HMI tags "Default tag table"
   "7" : Bool = PLC "ป้อนรหัส Barcode" AT %I100.6, 1 s
   "Alarms_All" : Word = PLC "บันทึกผลการเคลื่อนที่ ไว้ที่ Excell_DB".Alarms AT %DB1.DBX0.0, 1 s
   "Barcode1" : Word = PLC Barcode1 AT %MW2000, 1 s
   "Barcode10" : Word = PLC Barcode10 AT %MW2018, 1 s
   "Barcode100" : Word = PLC Barcode100 AT %MW2198, 1 s
   "Barcode101" : Word = PLC Barcode101 AT %MW2200, 1 s
   "Barcode102" : Word = PLC Barcode102 AT %MW2202, 1 s
   "Barcode103" : Word = PLC Barcode103 AT %MW2204, 1 s
   "Barcode104" : Word = PLC Barcode104 AT %MW2206, 1 s
   "Barcode105" : Word = PLC Barcode105 AT %MW2208, 1 s
   "Barcode106" : Word = PLC Barcode106 AT %MW2210, 1 s
   "Barcode107" : Word = PLC Barcode107 AT %MW2212, 1 s
   "Barcode108" : Word = PLC Barcode108 AT %MW2214, 1 s
   "Barcode109" : Word = PLC Barcode109 AT %MW2216, 1 s
   "Barcode11" : Word = PLC Barcode11 AT %MW2020, 1 s
   "Barcode110" : Word = PLC Barcode110 AT %MW2218, 1 s
   "Barcode111" : Word = PLC Barcode111 AT %MW2220, 1 s
   "Barcode112" : Word = PLC Barcode112 AT %MW2222, 1 s
   "Barcode113" : Word = PLC Barcode113 AT %MW2224, 1 s
   "Barcode114" : Word = PLC Barcode114 AT %MW2226, 1 s
   "Barcode115" : Word = PLC Barcode115 AT %MW2228, 1 s
   "Barcode116" : Word = PLC Barcode116 AT %MW2230, 1 s
   "Barcode117" : Word = PLC Barcode117 AT %MW2232, 1 s
   "Barcode118" : Word = PLC Barcode118 AT %MW2234, 1 s
   "Barcode119" : Word = PLC Barcode119 AT %MW2236, 1 s
   "Barcode12" : Word = PLC Barcode12 AT %MW2022, 1 s
   "Barcode120" : Word = PLC Barcode120 AT %MW2238, 1 s
   "Barcode121" : Word = PLC Barcode121 AT %MW2240, 1 s
   "Barcode122" : Word = PLC Barcode122 AT %MW2242, 1 s
   "Barcode123" : Word = PLC Barcode123 AT %MW2244, 1 s
   "Barcode124" : Word = PLC Barcode124 AT %MW2246, 1 s
   "Barcode125" : Word = PLC Barcode125 AT %MW2248, 1 s
   "Barcode126" : Word = PLC Barcode126 AT %MW2250, 1 s
   "Barcode127" : Word = PLC Barcode127 AT %MW2252, 1 s
   "Barcode128" : Word = PLC Barcode128 AT %MW2254, 1 s
   "Barcode129" : Word = PLC Barcode129 AT %MW2256, 1 s
   "Barcode13" : Word = PLC Barcode13 AT %MW2024, 1 s
   "Barcode130" : Word = PLC Barcode130 AT %MW2258, 1 s
   "Barcode131" : Word = PLC Barcode131 AT %MW2260, 1 s
   "Barcode132" : Word = PLC Barcode132 AT %MW2262, 1 s
   "Barcode133" : Word = PLC Barcode133 AT %MW2264, 1 s
   "Barcode134" : Word = PLC Barcode134 AT %MW2266, 1 s
   "Barcode135" : Word = PLC Barcode135 AT %MW2268, 1 s
   "Barcode136" : Word = PLC Barcode136 AT %MW2270, 1 s
   "Barcode137" : Word = PLC Barcode137 AT %MW2272, 1 s
   "Barcode138" : Word = PLC Barcode138 AT %MW2274, 1 s
   "Barcode139" : Word = PLC Barcode139 AT %MW2276, 1 s
   "Barcode14" : Word = PLC Barcode14 AT %MW2026, 1 s
   "Barcode140" : Word = PLC Barcode140 AT %MW2278, 1 s
   "Barcode141" : Word = PLC Barcode141 AT %MW2280, 1 s
   "Barcode142" : Word = PLC Barcode142 AT %MW2282, 1 s
   "Barcode143" : Word = PLC Barcode143 AT %MW2284, 1 s
   "Barcode144" : Word = PLC Barcode144 AT %MW2286, 1 s
   "Barcode145" : Word = PLC Barcode145 AT %MW2288, 1 s
   "Barcode146" : Word = PLC Barcode146 AT %MW2290, 1 s
   "Barcode147" : Word = PLC Barcode147 AT %MW2292, 1 s
   "Barcode148" : Word = PLC Barcode148 AT %MW2294, 1 s
   "Barcode149" : Word = PLC Barcode149 AT %MW2296, 1 s
   "Barcode15" : Word = PLC Barcode15 AT %MW2028, 1 s
   "Barcode150" : Word = PLC Barcode150 AT %MW2298, 1 s
   "Barcode151" : Word = PLC Barcode151 AT %MW2300, 1 s
   "Barcode152" : Word = PLC Barcode152 AT %MW2302, 1 s
   "Barcode153" : Word = PLC Barcode153 AT %MW2304, 1 s
   "Barcode154" : Word = PLC Barcode154 AT %MW2306, 1 s
   "Barcode155" : Word = PLC Barcode155 AT %MW2308, 1 s
   "Barcode156" : Word = PLC Barcode156 AT %MW2310, 1 s
   "Barcode157" : Word = PLC Barcode157 AT %MW2312, 1 s
   "Barcode158" : Word = PLC Barcode158 AT %MW2314, 1 s
   "Barcode159" : Word = PLC Barcode159 AT %MW2316, 1 s
   "Barcode16" : Word = PLC Barcode16 AT %MW2030, 1 s
   "Barcode160" : Word = PLC Barcode160 AT %MW2318, 1 s
   "Barcode161" : Word = PLC Barcode161 AT %MW2320, 1 s
   "Barcode162" : Word = PLC Barcode162 AT %MW2322, 1 s
   "Barcode163" : Word = PLC Barcode163 AT %MW2324, 1 s
   "Barcode164" : Word = PLC Barcode164 AT %MW2326, 1 s
   "Barcode165" : Word = PLC Barcode165 AT %MW2328, 1 s
   "Barcode166" : Word = PLC Barcode166 AT %MW2330, 1 s
   "Barcode167" : Word = PLC Barcode167 AT %MW2332, 1 s
   "Barcode168" : Word = PLC Barcode168 AT %MW2334, 1 s
   "Barcode169" : Word = PLC Barcode169 AT %MW2336, 1 s
   "Barcode17" : Word = PLC Barcode17 AT %MW2032, 1 s
   "Barcode170" : Word = PLC Barcode170 AT %MW2338, 1 s
   "Barcode171" : Word = PLC Barcode171 AT %MW2340, 1 s
   "Barcode172" : Word = PLC Barcode172 AT %MW2342, 1 s
   "Barcode173" : Word = PLC Barcode173 AT %MW2344, 1 s
   "Barcode174" : Word = PLC Barcode174 AT %MW2346, 1 s
   "Barcode175" : Word = PLC Barcode175 AT %MW2348, 1 s
   "Barcode176" : Word = PLC Barcode176 AT %MW2350, 1 s
   "Barcode177" : Word = PLC Barcode177 AT %MW2352, 1 s
   "Barcode178" : Word = PLC Barcode178 AT %MW2354, 1 s
   "Barcode179" : Word = PLC Barcode179 AT %MW2356, 1 s
   "Barcode18" : Word = PLC Barcode18 AT %MW2034, 1 s
   "Barcode180" : Word = PLC Barcode180 AT %MW2358, 1 s
   "Barcode181" : Word = PLC Barcode181 AT %MW2360, 1 s
   "Barcode182" : Word = PLC Barcode182 AT %MW2362, 1 s
   "Barcode183" : Word = PLC Barcode183 AT %MW2364, 1 s
   "Barcode184" : Word = PLC Barcode184 AT %MW2366, 1 s
   "Barcode185" : Word = PLC Barcode185 AT %MW2368, 1 s
   "Barcode186" : Word = PLC Barcode186 AT %MW2370, 1 s
   "Barcode187" : Word = PLC Barcode187 AT %MW2372, 1 s
   "Barcode188" : Word = PLC Barcode188 AT %MW2374, 1 s
   "Barcode189" : Word = PLC Barcode189 AT %MW2376, 1 s
   "Barcode19" : Word = PLC Barcode19 AT %MW2036, 1 s
   "Barcode190" : Word = PLC Barcode190 AT %MW2378, 1 s
   "Barcode191" : Word = PLC Barcode191 AT %MW2380, 1 s
   "Barcode192" : Word = PLC Barcode192 AT %MW2382, 1 s
   "Barcode193" : Word = PLC Barcode193 AT %MW2384, 1 s
   "Barcode194" : Word = PLC Barcode194 AT %MW2386, 1 s
   "Barcode195" : Word = PLC Barcode195 AT %MW2388, 1 s
   "Barcode196" : Word = PLC Barcode196 AT %MW2390, 1 s
   "Barcode197" : Word = PLC Barcode197 AT %MW2392, 1 s
   "Barcode198" : Word = PLC Barcode198 AT %MW2394, 1 s
   "Barcode199" : Word = PLC Barcode199 AT %MW2396, 1 s
   "Barcode2" : Word = PLC Barcode2 AT %MW2002, 1 s
   "Barcode20" : Word = PLC Barcode20 AT %MW2038, 1 s
   "Barcode200" : Word = PLC Barcode200 AT %MW2398, 1 s
   "Barcode201" : Word = PLC Barcode201 AT %MW2400, 1 s
   "Barcode202" : Word = PLC Barcode202 AT %MW2402, 1 s
   "Barcode203" : Word = PLC Barcode203 AT %MW2404, 1 s
   "Barcode204" : Word = PLC Barcode204 AT %MW2406, 1 s
   "Barcode205" : Word = PLC Barcode205 AT %MW2408, 1 s
   "Barcode206" : Word = PLC Barcode206 AT %MW2410, 1 s
   "Barcode207" : Word = PLC Barcode207 AT %MW2412, 1 s
   "Barcode208" : Word = PLC Barcode208 AT %MW2414, 1 s
   "Barcode209" : Word = PLC Barcode209 AT %MW2416, 1 s
   "Barcode21" : Word = PLC Barcode21 AT %MW2040, 1 s
   "Barcode210" : Word = PLC Barcode210 AT %MW2418, 1 s
   "Barcode211" : Word = PLC Barcode211 AT %MW2420, 1 s
   "Barcode212" : Word = PLC Barcode212 AT %MW2422, 1 s
   "Barcode213" : Word = PLC Barcode213 AT %MW2424, 1 s
   "Barcode214" : Word = PLC Barcode214 AT %MW2426, 1 s
   "Barcode215" : Word = PLC Barcode215 AT %MW2428, 1 s
   "Barcode216" : Word = PLC Barcode216 AT %MW2430, 1 s
   "Barcode217" : Word = PLC Barcode217 AT %MW2432, 1 s
   "Barcode218" : Word = PLC Barcode218 AT %MW2434, 1 s
   "Barcode219" : Word = PLC Barcode219 AT %MW2436, 1 s
   "Barcode22" : Word = PLC Barcode22 AT %MW2042, 1 s
   "Barcode220" : Word = PLC Barcode220 AT %MW2438, 1 s
   "Barcode221" : Word = PLC Barcode221 AT %MW2440, 1 s
   "Barcode222" : Word = PLC Barcode222 AT %MW2442, 1 s
   "Barcode223" : Word = PLC Barcode223 AT %MW2444, 1 s
   "Barcode224" : Word = PLC Barcode224 AT %MW2446, 1 s
   "Barcode225" : Word = PLC Barcode225 AT %MW2448, 1 s
   "Barcode226" : Word = PLC Barcode226 AT %MW2450, 1 s
   "Barcode227" : Word = PLC Barcode227 AT %MW2452, 1 s
   "Barcode228" : Word = PLC Barcode228 AT %MW2454, 1 s
   "Barcode229" : Word = PLC Barcode229 AT %MW2456, 1 s
   "Barcode23" : Word = PLC Barcode23 AT %MW2044, 1 s
   "Barcode230" : Word = PLC Barcode230 AT %MW2458, 1 s
   "Barcode231" : Word = PLC Barcode231 AT %MW2460, 1 s
   "Barcode232" : Word = PLC Barcode232 AT %MW2462, 1 s
   "Barcode233" : Word = PLC Barcode233 AT %MW2464, 1 s
   "Barcode234" : Word = PLC Barcode234 AT %MW2466, 1 s
   "Barcode235" : Word = PLC Barcode235 AT %MW2468, 1 s
   "Barcode236" : Word = PLC Barcode236 AT %MW2470, 1 s
   "Barcode237" : Word = PLC Barcode237 AT %MW2472, 1 s
   "Barcode238" : Word = PLC Barcode238 AT %MW2474, 1 s
   "Barcode239" : Word = PLC Barcode239 AT %MW2476, 1 s
   "Barcode24" : Word = PLC Barcode24 AT %MW2046, 1 s
   "Barcode240" : Word = PLC Barcode240 AT %MW2478, 1 s
   "Barcode241" : Word = PLC Barcode241 AT %MW2480, 1 s
   "Barcode242" : Word = PLC Barcode242 AT %MW2482, 1 s
   "Barcode243" : Word = PLC Barcode243 AT %MW2484, 1 s
   "Barcode244" : Word = PLC Barcode244 AT %MW2486, 1 s
   "Barcode245" : Word = PLC Barcode245 AT %MW2488, 1 s
   "Barcode246" : Word = PLC Barcode246 AT %MW2490, 1 s
   "Barcode247" : Word = PLC Barcode247 AT %MW2492, 1 s
   "Barcode248" : Word = PLC Barcode248 AT %MW2494, 1 s
   "Barcode249" : Word = PLC Barcode249 AT %MW2496, 1 s
   "Barcode25" : Word = PLC Barcode25 AT %MW2048, 1 s
   "Barcode250" : Word = PLC Barcode250 AT %MW2498, 1 s
   "Barcode251" : Word = PLC Barcode251 AT %MW2500, 1 s
   "Barcode252" : Word = PLC Barcode252 AT %MW2502, 1 s
   "Barcode253" : Word = PLC Barcode253 AT %MW2504, 1 s
   "Barcode254" : Word = PLC Barcode254 AT %MW2506, 1 s
   "Barcode255" : Word = PLC Barcode255 AT %MW2508, 1 s
   "Barcode256" : Word = PLC Barcode256 AT %MW2510, 1 s
   "Barcode257" : Word = PLC Barcode257 AT %MW2512, 1 s
   "Barcode258" : Word = PLC Barcode258 AT %MW2514, 1 s
   "Barcode259" : Word = PLC Barcode259 AT %MW2516, 1 s
   "Barcode26" : Word = PLC Barcode26 AT %MW2050, 1 s
   "Barcode260" : Word = PLC Barcode260 AT %MW2518, 1 s
   "Barcode261" : Word = PLC Barcode261 AT %MW2520, 1 s
   "Barcode262" : Word = PLC Barcode262 AT %MW2522, 1 s
   "Barcode263" : Word = PLC Barcode263 AT %MW2524, 1 s
   "Barcode264" : Word = PLC Barcode264 AT %MW2526, 1 s
   "Barcode265" : Word = PLC Barcode265 AT %MW2528, 1 s
   "Barcode266" : Word = PLC Barcode266 AT %MW2530, 1 s
   "Barcode267" : Word = PLC Barcode267 AT %MW2532, 1 s
   "Barcode268" : Word = PLC Barcode268 AT %MW2534, 1 s
   "Barcode269" : Word = PLC Barcode269 AT %MW2536, 1 s
   "Barcode27" : Word = PLC Barcode27 AT %MW2052, 1 s
   "Barcode270" : Word = PLC Barcode270 AT %MW2538, 1 s
   "Barcode271" : Word = PLC Barcode271 AT %MW2540, 1 s
   "Barcode272" : Word = PLC Barcode272 AT %MW2542, 1 s
   "Barcode273" : Word = PLC Barcode273 AT %MW2544, 1 s
   "Barcode274" : Word = PLC Barcode274 AT %MW2546, 1 s
   "Barcode275" : Word = PLC Barcode275 AT %MW2548, 1 s
   "Barcode276" : Word = PLC Barcode276 AT %MW2550, 1 s
   "Barcode277" : Word = PLC Barcode277 AT %MW2552, 1 s
   "Barcode278" : Word = PLC Barcode278 AT %MW2554, 1 s
   "Barcode279" : Word = PLC Barcode279 AT %MW2556, 1 s
   "Barcode28" : Word = PLC Barcode28 AT %MW2054, 1 s
   "Barcode280" : Word = PLC Barcode280 AT %MW2558, 1 s
   "Barcode281" : Word = PLC Barcode281 AT %MW2560, 1 s
   "Barcode282" : Word = PLC Barcode282 AT %MW2562, 1 s
   "Barcode283" : Word = PLC Barcode283 AT %MW2564, 1 s
   "Barcode284" : Word = PLC Barcode284 AT %MW2566, 1 s
   "Barcode285" : Word = PLC Barcode285 AT %MW2568, 1 s
   "Barcode286" : Word = PLC Barcode286 AT %MW2570, 1 s
   "Barcode287" : Word = PLC Barcode287 AT %MW2572, 1 s
   "Barcode288" : Word = PLC Barcode288 AT %MW2574, 1 s
   "Barcode289" : Word = PLC Barcode289 AT %MW2576, 1 s
   "Barcode29" : Word = PLC Barcode29 AT %MW2056, 1 s
   "Barcode290" : Word = PLC Barcode290 AT %MW2578, 1 s
   "Barcode291" : Word = PLC Barcode291 AT %MW2580, 1 s
   "Barcode292" : Word = PLC Barcode292 AT %MW2582, 1 s
   "Barcode293" : Word = PLC Barcode293 AT %MW2584, 1 s
   "Barcode294" : Word = PLC Barcode294 AT %MW2586, 1 s
   "Barcode295" : Word = PLC Barcode295 AT %MW2588, 1 s
   "Barcode296" : Word = PLC Barcode296 AT %MW2590, 1 s
   "Barcode297" : Word = PLC Barcode297 AT %MW2592, 1 s
   "Barcode298" : Word = PLC Barcode298 AT %MW2594, 1 s
   "Barcode299" : Word = PLC Barcode299 AT %MW2596, 1 s
   "Barcode3" : Word = PLC Barcode3 AT %MW2004, 1 s
   "Barcode30" : Word = PLC Barcode30 AT %MW2058, 1 s
   "Barcode300" : Word = PLC Barcode300 AT %MW2598, 1 s
   "Barcode301" : Word = PLC Barcode301 AT %MW2600, 1 s
   "Barcode302" : Word = PLC Barcode302 AT %MW2602, 1 s
   "Barcode303" : Word = PLC Barcode303 AT %MW2604, 1 s
   "Barcode304" : Word = PLC Barcode304 AT %MW2606, 1 s
   "Barcode305" : Word = PLC Barcode305 AT %MW2608, 1 s
   "Barcode306" : Word = PLC Barcode306 AT %MW2610, 1 s
   "Barcode307" : Word = PLC Barcode307 AT %MW2612, 1 s
   "Barcode308" : Word = PLC Barcode308 AT %MW2614, 1 s
   "Barcode309" : Word = PLC Barcode309 AT %MW2616, 1 s
   "Barcode31" : Word = PLC Barcode31 AT %MW2060, 1 s
   "Barcode310" : Word = PLC Barcode310 AT %MW2618, 1 s
   "Barcode311" : Word = PLC Barcode311 AT %MW2620, 1 s
   "Barcode312" : Word = PLC Barcode312 AT %MW2622, 1 s
   "Barcode313" : Word = PLC Barcode313 AT %MW2624, 1 s
   "Barcode314" : Word = PLC Barcode314 AT %MW2626, 1 s
   "Barcode315" : Word = PLC Barcode315 AT %MW2628, 1 s
   "Barcode316" : Word = PLC Barcode316 AT %MW2630, 1 s
   "Barcode317" : Word = PLC Barcode317 AT %MW2632, 1 s
   "Barcode318" : Word = PLC Barcode318 AT %MW2634, 1 s
   "Barcode319" : Word = PLC Barcode319 AT %MW2636, 1 s
   "Barcode32" : Word = PLC Barcode32 AT %MW2062, 1 s
   "Barcode320" : Word = PLC Barcode320 AT %MW2638, 1 s
   "Barcode321" : Word = PLC Barcode321 AT %MW2640, 1 s
   "Barcode322" : Word = PLC Barcode322 AT %MW2642, 1 s
   "Barcode323" : Word = PLC Barcode323 AT %MW2644, 1 s
   "Barcode324" : Word = PLC Barcode324 AT %MW2646, 1 s
   "Barcode325" : Word = PLC Barcode325 AT %MW2648, 1 s
   "Barcode326" : Word = PLC Barcode326 AT %MW2650, 1 s
   "Barcode327" : Word = PLC Barcode327 AT %MW2652, 1 s
   "Barcode328" : Word = PLC Barcode328 AT %MW2654, 1 s
   "Barcode329" : Word = PLC Barcode329 AT %MW2656, 1 s
   "Barcode33" : Word = PLC Barcode33 AT %MW2064, 1 s
   "Barcode330" : Word = PLC Barcode330 AT %MW2658, 1 s
   "Barcode331" : Word = PLC Barcode331 AT %MW2660, 1 s
   "Barcode332" : Word = PLC Barcode332 AT %MW2662, 1 s
   "Barcode333" : Word = PLC Barcode333 AT %MW2664, 1 s
   "Barcode334" : Word = PLC Barcode334 AT %MW2666, 1 s
   "Barcode335" : Word = PLC Barcode335 AT %MW2668, 1 s
   "Barcode336" : Word = PLC Barcode336 AT %MW2670, 1 s
   "Barcode337" : Word = PLC Barcode337 AT %MW2672, 1 s
   "Barcode338" : Word = PLC Barcode338 AT %MW2674, 1 s
   "Barcode339" : Word = PLC Barcode339 AT %MW2676, 1 s
   "Barcode34" : Word = PLC Barcode34 AT %MW2066, 1 s
   "Barcode340" : Word = PLC Barcode340 AT %MW2678, 1 s
   "Barcode341" : Word = PLC Barcode341 AT %MW2680, 1 s
   "Barcode342" : Word = PLC Barcode342 AT %MW2682, 1 s
   "Barcode343" : Word = PLC Barcode343 AT %MW2684, 1 s
   "Barcode344" : Word = PLC Barcode344 AT %MW2686, 1 s
   "Barcode345" : Word = PLC Barcode345 AT %MW2688, 1 s
   "Barcode346" : Word = PLC Barcode346 AT %MW2690, 1 s
   "Barcode347" : Word = PLC Barcode347 AT %MW2692, 1 s
   "Barcode348" : Word = PLC Barcode348 AT %MW2694, 1 s
   "Barcode349" : Word = PLC Barcode349 AT %MW2696, 1 s
   "Barcode35" : Word = PLC Barcode35 AT %MW2068, 1 s
   "Barcode350" : Word = PLC Barcode350 AT %MW2698, 1 s
   "Barcode351" : Word = PLC Barcode351 AT %MW2700, 1 s
   "Barcode352" : Word = PLC Barcode352 AT %MW2702, 1 s
   "Barcode353" : Word = PLC Barcode353 AT %MW2704, 1 s
   "Barcode354" : Word = PLC Barcode354 AT %MW2706, 1 s
   "Barcode355" : Word = PLC Barcode355 AT %MW2708, 1 s
   "Barcode356" : Word = PLC Barcode356 AT %MW2710, 1 s
   "Barcode357" : Word = PLC Barcode357 AT %MW2712, 1 s
   "Barcode358" : Word = PLC Barcode358 AT %MW2714, 1 s
   "Barcode359" : Word = PLC Barcode359 AT %MW2716, 1 s
   "Barcode36" : Word = PLC Barcode36 AT %MW2070, 1 s
   "Barcode360" : Word = PLC Barcode360 AT %MW2718, 1 s
   "Barcode361" : Word = PLC Barcode361 AT %MW2720, 1 s
   "Barcode362" : Word = PLC Barcode362 AT %MW2722, 1 s
   "Barcode363" : Word = PLC Barcode363 AT %MW2724, 1 s
   "Barcode364" : Word = PLC Barcode364 AT %MW2726, 1 s
   "Barcode365" : Word = PLC Barcode365 AT %MW2728, 1 s
   "Barcode366" : Word = PLC Barcode366 AT %MW2730, 1 s
   "Barcode367" : Word = PLC Barcode367 AT %MW2732, 1 s
   "Barcode368" : Word = PLC Barcode368 AT %MW2734, 1 s
   "Barcode369" : Word = PLC Barcode369 AT %MW2736, 1 s
   "Barcode37" : Word = PLC Barcode37 AT %MW2072, 1 s
   "Barcode370" : Word = PLC Barcode370 AT %MW2738, 1 s
   "Barcode371" : Word = PLC Barcode371 AT %MW2740, 1 s
   "Barcode372" : Word = PLC Barcode372 AT %MW2742, 1 s
   "Barcode373" : Word = PLC Barcode373 AT %MW2744, 1 s
   "Barcode374" : Word = PLC Barcode374 AT %MW2746, 1 s
   "Barcode375" : Word = PLC Barcode375 AT %MW2748, 1 s
   "Barcode376" : Word = PLC Barcode376 AT %MW2750, 1 s
   "Barcode377" : Word = PLC Barcode377 AT %MW2752, 1 s
   "Barcode378" : Word = PLC Barcode378 AT %MW2754, 1 s
   "Barcode379" : Word = PLC Barcode379 AT %MW2756, 1 s
   "Barcode38" : Word = PLC Barcode38 AT %MW2074, 1 s
   "Barcode380" : Word = PLC Barcode380 AT %MW2758, 1 s
   "Barcode381" : Word = PLC Barcode381 AT %MW2760, 1 s
   "Barcode382" : Word = PLC Barcode382 AT %MW2762, 1 s
   "Barcode383" : Word = PLC Barcode383 AT %MW2764, 1 s
   "Barcode384" : Word = PLC Barcode384 AT %MW2766, 1 s
   "Barcode385" : Word = PLC Barcode385 AT %MW2768, 1 s
   "Barcode386" : Word = PLC Barcode386 AT %MW2770, 1 s
   "Barcode387" : Word = PLC Barcode387 AT %MW2772, 1 s
   "Barcode388" : Word = PLC Barcode388 AT %MW2774, 1 s
   "Barcode389" : Word = PLC Barcode389 AT %MW2776, 1 s
   "Barcode39" : Word = PLC Barcode39 AT %MW2076, 1 s
   "Barcode390" : Word = PLC Barcode390 AT %MW2778, 1 s
   "Barcode391" : Word = PLC Barcode391 AT %MW2780, 1 s
   "Barcode392" : Word = PLC Barcode392 AT %MW2782, 1 s
   "Barcode393" : Word = PLC Barcode393 AT %MW2784, 1 s
   "Barcode394" : Word = PLC Barcode394 AT %MW2786, 1 s
   "Barcode395" : Word = PLC Barcode395 AT %MW2788, 1 s
   "Barcode396" : Word = PLC Barcode396 AT %MW2790, 1 s
   "Barcode397" : Word = PLC Barcode397 AT %MW2792, 1 s
   "Barcode398" : Word = PLC Barcode398 AT %MW2794, 1 s
   "Barcode399" : Word = PLC Barcode399 AT %MW2796, 1 s
   "Barcode4" : Word = PLC Barcode4 AT %MW2006, 1 s
   "Barcode40" : Word = PLC Barcode40 AT %MW2078, 1 s
   "Barcode400" : Word = PLC Barcode400 AT %MW2798, 1 s
   "Barcode401" : Word = PLC Barcode401 AT %MW2800, 1 s
   "Barcode402" : Word = PLC Barcode402 AT %MW2802, 1 s
   "Barcode403" : Word = PLC Barcode403 AT %MW2804, 1 s
   "Barcode404" : Word = PLC Barcode404 AT %MW2806, 1 s
   "Barcode405" : Word = PLC Barcode405 AT %MW2808, 1 s
   "Barcode406" : Word = PLC Barcode406 AT %MW2810, 1 s
   "Barcode407" : Word = PLC Barcode407 AT %MW2812, 1 s
   "Barcode408" : Word = PLC Barcode408 AT %MW2814, 1 s
   "Barcode409" : Word = PLC Barcode409 AT %MW2816, 1 s
   "Barcode41" : Word = PLC Barcode41 AT %MW2080, 1 s
   "Barcode410" : Word = PLC Barcode410 AT %MW2818, 1 s
   "Barcode411" : Word = PLC Barcode411 AT %MW2820, 1 s
   "Barcode412" : Word = PLC Barcode412 AT %MW2822, 1 s
   "Barcode413" : Word = PLC Barcode413 AT %MW2824, 1 s
   "Barcode414" : Word = PLC Barcode414 AT %MW2826, 1 s
   "Barcode415" : Word = PLC Barcode415 AT %MW2828, 1 s
   "Barcode416" : Word = PLC Barcode416 AT %MW2830, 1 s
   "Barcode417" : Word = PLC Barcode417 AT %MW2832, 1 s
   "Barcode418" : Word = PLC Barcode418 AT %MW2834, 1 s
   "Barcode419" : Word = PLC Barcode419 AT %MW2836, 1 s
   "Barcode42" : Word = PLC Barcode42 AT %MW2082, 1 s
   "Barcode420" : Word = PLC Barcode420 AT %MW2838, 1 s
   "Barcode421" : Word = PLC Barcode421 AT %MW2840, 1 s
   "Barcode422" : Word = PLC Barcode422 AT %MW2842, 1 s
   "Barcode423" : Word = PLC Barcode423 AT %MW2844, 1 s
   "Barcode424" : Word = PLC Barcode424 AT %MW2846, 1 s
   "Barcode425" : Word = PLC Barcode425 AT %MW2848, 1 s
   "Barcode426" : Word = PLC Barcode426 AT %MW2850, 1 s
   "Barcode427" : Word = PLC Barcode427 AT %MW2852, 1 s
   "Barcode428" : Word = PLC Barcode428 AT %MW2854, 1 s
   "Barcode429" : Word = PLC Barcode429 AT %MW2856, 1 s
   "Barcode43" : Word = PLC Barcode43 AT %MW2084, 1 s
   "Barcode430" : Word = PLC Barcode430 AT %MW2858, 1 s
   "Barcode431" : Word = PLC Barcode431 AT %MW2860, 1 s
   "Barcode432" : Word = PLC Barcode432 AT %MW2862, 1 s
   "Barcode433" : Word = PLC Barcode433 AT %MW2864, 1 s
   "Barcode434" : Word = PLC Barcode434 AT %MW2866, 1 s
   "Barcode435" : Word = PLC Barcode435 AT %MW2868, 1 s
   "Barcode436" : Word = PLC Barcode436 AT %MW2870, 1 s
   "Barcode437" : Word = PLC Barcode437 AT %MW2872, 1 s
   "Barcode438" : Word = PLC Barcode438 AT %MW2874, 1 s
   "Barcode439" : Word = PLC Barcode439 AT %MW2876, 1 s
   "Barcode44" : Word = PLC Barcode44 AT %MW2086, 1 s
   "Barcode440" : Word = PLC Barcode440 AT %MW2878, 1 s
   "Barcode441" : Word = PLC Barcode441 AT %MW2880, 1 s
   "Barcode442" : Word = PLC Barcode442 AT %MW2882, 1 s
   "Barcode443" : Word = PLC Barcode443 AT %MW2884, 1 s
   "Barcode444" : Word = PLC Barcode444 AT %MW2886, 1 s
   "Barcode445" : Word = PLC Barcode445 AT %MW2888, 1 s
   "Barcode446" : Word = PLC Barcode446 AT %MW2890, 1 s
   "Barcode447" : Word = PLC Barcode447 AT %MW2892, 1 s
   "Barcode448" : Word = PLC Barcode448 AT %MW2894, 1 s
   "Barcode449" : Word = PLC Barcode449 AT %MW2896, 1 s
   "Barcode45" : Word = PLC Barcode45 AT %MW2088, 1 s
   "Barcode450" : Word = PLC Barcode450 AT %MW2898, 1 s
   "Barcode451" : Word = PLC Barcode451 AT %MW2900, 1 s
   "Barcode452" : Word = PLC Barcode452 AT %MW2902, 1 s
   "Barcode453" : Word = PLC Barcode453 AT %MW2904, 1 s
   "Barcode454" : Word = PLC Barcode454 AT %MW2906, 1 s
   "Barcode455" : Word = PLC Barcode455 AT %MW2908, 1 s
   "Barcode456" : Word = PLC Barcode456 AT %MW2910, 1 s
   "Barcode457" : Word = PLC Barcode457 AT %MW2912, 1 s
   "Barcode458" : Word = PLC Barcode458 AT %MW2914, 1 s
   "Barcode459" : Word = PLC Barcode459 AT %MW2916, 1 s
   "Barcode46" : Word = PLC Barcode46 AT %MW2090, 1 s
   "Barcode460" : Word = PLC Barcode460 AT %MW2918, 1 s
   "Barcode461" : Word = PLC Barcode461 AT %MW2920, 1 s
   "Barcode462" : Word = PLC Barcode462 AT %MW2922, 1 s
   "Barcode463" : Word = PLC Barcode463 AT %MW2924, 1 s
   "Barcode464" : Word = PLC Barcode464 AT %MW2926, 1 s
   "Barcode465" : Word = PLC Barcode465 AT %MW2928, 1 s
   "Barcode466" : Word = PLC Barcode466 AT %MW2930, 1 s
   "Barcode467" : Word = PLC Barcode467 AT %MW2932, 1 s
   "Barcode468" : Word = PLC Barcode468 AT %MW2934, 1 s
   "Barcode469" : Word = PLC Barcode469 AT %MW2936, 1 s
   "Barcode47" : Word = PLC Barcode47 AT %MW2092, 1 s
   "Barcode470" : Word = PLC Barcode470 AT %MW2938, 1 s
   "Barcode471" : Word = PLC Barcode471 AT %MW2940, 1 s
   "Barcode472" : Word = PLC Barcode472 AT %MW2942, 1 s
   "Barcode473" : Word = PLC Barcode473 AT %MW2944, 1 s
   "Barcode474" : Word = PLC Barcode474 AT %MW2946, 1 s
   "Barcode475" : Word = PLC Barcode475 AT %MW2948, 1 s
   "Barcode476" : Word = PLC Barcode476 AT %MW2950, 1 s
   "Barcode477" : Word = PLC Barcode477 AT %MW2952, 1 s
   "Barcode478" : Word = PLC Barcode478 AT %MW2954, 1 s
   "Barcode479" : Word = PLC Barcode479 AT %MW2956, 1 s
   "Barcode48" : Word = PLC Barcode48 AT %MW2094, 1 s
   "Barcode480" : Word = PLC Barcode480 AT %MW2958, 1 s
   "Barcode481" : Word = PLC Barcode481 AT %MW2960, 1 s
   "Barcode482" : Word = PLC Barcode482 AT %MW2962, 1 s
   "Barcode483" : Word = PLC Barcode483 AT %MW2964, 1 s
   "Barcode484" : Word = PLC Barcode484 AT %MW2966, 1 s
   "Barcode485" : Word = PLC Barcode485 AT %MW2968, 1 s
   "Barcode486" : Word = PLC Barcode486 AT %MW2970, 1 s
   "Barcode487" : Word = PLC Barcode487 AT %MW2972, 1 s
   "Barcode488" : Word = PLC Barcode488 AT %MW2974, 1 s
   "Barcode489" : Word = PLC Barcode489 AT %MW2976, 1 s
   "Barcode49" : Word = PLC Barcode49 AT %MW2096, 1 s
   "Barcode490" : Word = PLC Barcode490 AT %MW2978, 1 s
   "Barcode491" : Word = PLC Barcode491 AT %MW2980, 1 s
   "Barcode492" : Word = PLC Barcode492 AT %MW2982, 1 s
   "Barcode493" : Word = PLC Barcode493 AT %MW2984, 1 s
   "Barcode494" : Word = PLC Barcode494 AT %MW2986, 1 s
   "Barcode495" : Word = PLC Barcode495 AT %MW2988, 1 s
   "Barcode496" : Word = PLC Barcode496 AT %MW2990, 1 s
   "Barcode497" : Word = PLC Barcode497 AT %MW2992, 1 s
   "Barcode498" : Word = PLC Barcode498 AT %MW2994, 1 s
   "Barcode499" : Word = PLC Barcode499 AT %MW2996, 1 s
   "Barcode5" : Word = PLC Barcode5 AT %MW2008, 1 s
   "Barcode50" : Word = PLC Barcode50 AT %MW2098, 1 s
   "Barcode500" : Word = PLC Barcode500 AT %MW2998, 1 s
   "Barcode501" : Word = PLC Barcode501 AT %MW3000, 1 s
   "Barcode502" : Word = PLC Barcode502 AT %MW3002, 1 s
   "Barcode503" : Word = PLC Barcode503 AT %MW3004, 1 s
   "Barcode504" : Word = PLC Barcode504 AT %MW3006, 1 s
   "Barcode505" : Word = PLC Barcode505 AT %MW3008, 1 s
   "Barcode506" : Word = PLC Barcode506 AT %MW3010, 1 s
   "Barcode507" : Word = PLC Barcode507 AT %MW3012, 1 s
   "Barcode508" : Word = PLC Barcode508 AT %MW3014, 1 s
   "Barcode509" : Word = PLC Barcode509 AT %MW3016, 1 s
   "Barcode51" : Word = PLC Barcode51 AT %MW2100, 1 s
   "Barcode510" : Word = PLC Barcode510 AT %MW3018, 1 s
   "Barcode511" : Word = PLC Barcode511 AT %MW3020, 1 s
   "Barcode512" : Word = PLC Barcode512 AT %MW3022, 1 s
   "Barcode513" : Word = PLC Barcode513 AT %MW3024, 1 s
   "Barcode514" : Word = PLC Barcode514 AT %MW3026, 1 s
   "Barcode515" : Word = PLC Barcode515 AT %MW3028, 1 s
   "Barcode516" : Word = PLC Barcode516 AT %MW3030, 1 s
   "Barcode517" : Word = PLC Barcode517 AT %MW3032, 1 s
   "Barcode518" : Word = PLC Barcode518 AT %MW3034, 1 s
   "Barcode519" : Word = PLC Barcode519 AT %MW3036, 1 s
   "Barcode52" : Word = PLC Barcode52 AT %MW2102, 1 s
   "Barcode520" : Word = PLC Barcode520 AT %MW3038, 1 s
   "Barcode53" : Word = PLC Barcode53 AT %MW2104, 1 s
   "Barcode54" : Word = PLC Barcode54 AT %MW2106, 1 s
   "Barcode55" : Word = PLC Barcode55 AT %MW2108, 1 s
   "Barcode56" : Word = PLC Barcode56 AT %MW2110, 1 s
   "Barcode57" : Word = PLC Barcode57 AT %MW2112, 1 s
   "Barcode58" : Word = PLC Barcode58 AT %MW2114, 1 s
   "Barcode59" : Word = PLC Barcode59 AT %MW2116, 1 s
   "Barcode6" : Word = PLC Barcode6 AT %MW2010, 1 s
   "Barcode60" : Word = PLC Barcode60 AT %MW2118, 1 s
   "Barcode61" : Word = PLC Barcode61 AT %MW2120, 1 s
   "Barcode62" : Word = PLC Barcode62 AT %MW2122, 1 s
   "Barcode63" : Word = PLC Barcode63 AT %MW2124, 1 s
   "Barcode64" : Word = PLC Barcode64 AT %MW2126, 1 s
   "Barcode65" : Word = PLC Barcode65 AT %MW2128, 1 s
   "Barcode66" : Word = PLC Barcode66 AT %MW2130, 1 s
   "Barcode67" : Word = PLC Barcode67 AT %MW2132, 1 s
   "Barcode68" : Word = PLC Barcode68 AT %MW2134, 1 s
   "Barcode69" : Word = PLC Barcode69 AT %MW2136, 1 s
   "Barcode7" : Word = PLC Barcode7 AT %MW2012, 1 s
   "Barcode70" : Word = PLC Barcode70 AT %MW2138, 1 s
   "Barcode71" : Word = PLC Barcode71 AT %MW2140, 1 s
   "Barcode72" : Word = PLC Barcode72 AT %MW2142, 1 s
   "Barcode73" : Word = PLC Barcode73 AT %MW2144, 1 s
   "Barcode74" : Word = PLC Barcode74 AT %MW2146, 1 s
   "Barcode75" : Word = PLC Barcode75 AT %MW2148, 1 s
   "Barcode76" : Word = PLC Barcode76 AT %MW2150, 1 s
   "Barcode77" : Word = PLC Barcode77 AT %MW2152, 1 s
   "Barcode78" : Word = PLC Barcode78 AT %MW2154, 1 s
   "Barcode79" : Word = PLC Barcode79 AT %MW2156, 1 s
   "Barcode8" : Word = PLC Barcode8 AT %MW2014, 1 s
   "Barcode80" : Word = PLC Barcode80 AT %MW2158, 1 s
   "Barcode81" : Word = PLC Barcode81 AT %MW2160, 1 s
   "Barcode82" : Word = PLC Barcode82 AT %MW2162, 1 s
   "Barcode83" : Word = PLC Barcode83 AT %MW2164, 1 s
   "Barcode84" : Word = PLC Barcode84 AT %MW2166, 1 s
   "Barcode85" : Word = PLC Barcode85 AT %MW2168, 1 s
   "Barcode86" : Word = PLC Barcode86 AT %MW2170, 1 s
   "Barcode87" : Word = PLC Barcode87 AT %MW2172, 1 s
   "Barcode88" : Word = PLC Barcode88 AT %MW2174, 1 s
   "Barcode89" : Word = PLC Barcode89 AT %MW2176, 1 s
   "Barcode9" : Word = PLC Barcode9 AT %MW2016, 1 s
   "Barcode90" : Word = PLC Barcode90 AT %MW2178, 1 s
   "Barcode91" : Word = PLC Barcode91 AT %MW2180, 1 s
   "Barcode92" : Word = PLC Barcode92 AT %MW2182, 1 s
   "Barcode93" : Word = PLC Barcode93 AT %MW2184, 1 s
   "Barcode94" : Word = PLC Barcode94 AT %MW2186, 1 s
   "Barcode95" : Word = PLC Barcode95 AT %MW2188, 1 s
   "Barcode96" : Word = PLC Barcode96 AT %MW2190, 1 s
   "Barcode97" : Word = PLC Barcode97 AT %MW2192, 1 s
   "Barcode98" : Word = PLC Barcode98 AT %MW2194, 1 s
   "Barcode99" : Word = PLC Barcode99 AT %MW2196, 1 s
   "Button_OK_Screen" : Bool = PLC Button_OK_Screen AT %M3040.0, 1 s
   "Expected/Value_All_V" : String[254] = PLC "Expected/Value_All".V, 1 s
   "Gripper เคลื่อนไปช่องยา" : Bool = PLC "Gripper เคลื่อนไปช่องยา" AT %I101.0, 1 s
   "Gripper วางยา" : Bool = PLC "Gripper วางยา" AT %I101.1, 1 s
   "Gripper หยิบยา" : Bool = PLC "Gripper หยิบยา" AT %I102.1, 1 s
   "Gripperเคลื่อนที่มาเอายา" : Bool = PLC Gripperเคลื่อนที่มาเอายา AT %I100.7, 1 s
   "Output Status1" : Word = PLC "Output Status1" AT %MW3054, 1 s
   "Output Status2" : Word = PLC "Output Status2" AT %MW3056, 1 s
   "Selected_Medicine" : Int AT %DB1.DBW0
   "Selected_Medicine_final" : Int AT %DB1.DBX0.0
   "Selected_URL" : WString[254], internal
   "Video_URL" : WString[254] AT %DB1.DBX0.0
   "เคลื่อนที่ไปยังจุดเริ่มต้น" : Bool = PLC เคลื่อนที่ไปยังจุดเริ่มต้น AT %I101.2, 1 s
   "เคลื่อนที่ไปยังตำแหน่งเริ่มต้น เบิกจ่าย" : Bool = PLC "เคลื่อนที่ไปยังตำแหน่งเริ่มต้น เบิกจ่าย" AT %I101.7, 1 s
   "เคลื่อนที่ไปยังตำยา" : Bool = PLC เคลื่อนที่ไปยังตำยา AT %I101.5, 1 s
   "เบิกจ่าย Servo DATA 1,2" : Word = PLC "เบิกจ่าย Servo DATA 1,2" AT %MW3050, 1 s
   "เบิกจ่าย Servo DATA 3" : Word = PLC "เบิกจ่าย Servo DATA 3" AT %MW3052, 1 s
   "แสดงชื่อยา" : Word = PLC แสดงชื่อยา AT %MW3042, 1 s
   "แสดงชื่อยา2" : Word = PLC แสดงชื่อยา2 AT %MW3044, 1 s
   "จัดเก็บ Servo DATA 1,2" : Word = PLC "จัดเก็บ Servo DATA 1,2" AT %MW3046, 1 s
   "จัดเก็บ Servo DATA 3" : Word = PLC "จัดเก็บ Servo DATA 3" AT %MW3048, 1 s
   "ป้อนรหัส Barcode" : Bool = PLC "ป้อนรหัส Barcode" AT %I100.6, 1 s
   "ปุ่มClear" : Bool = PLC ปุ่มClear AT %M1965.2, 1 s
   "ปุ่มยืนยันหน้า Screen" : Bool = PLC "ปุ่มยืนยันหน้า Screen" AT %M1965.0, 1 s
   "มีการปุ่มกดยืนยัน" : Bool = PLC มีการปุ่มกดยืนยัน AT %M100.2, 1 s
   "ยา 1" : Word = PLC "ยา 1" AT %MW850, 1 s
   "ยา 10" : Word = PLC "ยา 10" AT %MW868, 1 s
   "ยา 100" : Word = PLC "ยา 100" AT %MW1048, 1 s
   "ยา 101" : Word = PLC "ยา 101" AT %MW1050, 1 s
   "ยา 102" : Word = PLC "ยา 102" AT %MW1052, 1 s
   "ยา 103" : Word = PLC "ยา 103" AT %MW1054, 1 s
   "ยา 104" : Word = PLC "ยา 104" AT %MW1056, 1 s
   "ยา 105" : Word = PLC "ยา 105" AT %MW1058, 1 s
   "ยา 106" : Word = PLC "ยา 106" AT %MW1060, 1 s
   "ยา 107" : Word = PLC "ยา 107" AT %MW1062, 1 s
   "ยา 108" : Word = PLC "ยา 108" AT %MW1064, 1 s
   "ยา 109" : Word = PLC "ยา 109" AT %MW1066, 1 s
   "ยา 11" : Word = PLC "ยา 11" AT %MW870, 1 s
   "ยา 110" : Word = PLC "ยา 110" AT %MW1068, 1 s
   "ยา 111" : Word = PLC "ยา 111" AT %MW1070, 1 s
   "ยา 112" : Word = PLC "ยา 112" AT %MW1072, 1 s
   "ยา 113" : Word = PLC "ยา 113" AT %MW1074, 1 s
   "ยา 114" : Word = PLC "ยา 114" AT %MW1076, 1 s
   "ยา 115" : Word = PLC "ยา 115" AT %MW1078, 1 s
   "ยา 116" : Word = PLC "ยา 116" AT %MW1080, 1 s
   "ยา 117" : Word = PLC "ยา 117" AT %MW1082, 1 s
   "ยา 118" : Word = PLC "ยา 118" AT %MW1084, 1 s
   "ยา 119" : Word = PLC "ยา 119" AT %MW1086, 1 s
   "ยา 12" : Word = PLC "ยา 12" AT %MW872, 1 s
   "ยา 120" : Word = PLC "ยา 120" AT %MW1088, 1 s
   "ยา 121" : Word = PLC "ยา 121" AT %MW1090, 1 s
   "ยา 122" : Word = PLC "ยา 122" AT %MW1092, 1 s
   "ยา 123" : Word = PLC "ยา 123" AT %MW1094, 1 s
   "ยา 124" : Word = PLC "ยา 124" AT %MW1096, 1 s
   "ยา 125" : Word = PLC "ยา 125" AT %MW1098, 1 s
   "ยา 126" : Word = PLC "ยา 126" AT %MW1100, 1 s
   "ยา 127" : Word = PLC "ยา 127" AT %MW1102, 1 s
   "ยา 128" : Word = PLC "ยา 128" AT %MW1104, 1 s
   "ยา 129" : Word = PLC "ยา 129" AT %MW1106, 1 s
   "ยา 13" : Word = PLC "ยา 13" AT %MW874, 1 s
   "ยา 130" : Word = PLC "ยา 130" AT %MW1108, 1 s
   "ยา 131" : Word = PLC "ยา 131" AT %MW1110, 1 s
   "ยา 132" : Word = PLC "ยา 132" AT %MW1112, 1 s
   "ยา 133" : Word = PLC "ยา 133" AT %MW1114, 1 s
   "ยา 134" : Word = PLC "ยา 134" AT %MW1116, 1 s
   "ยา 135" : Word = PLC "ยา 135" AT %MW1118, 1 s
   "ยา 136" : Word = PLC "ยา 136" AT %MW1120, 1 s
   "ยา 137" : Word = PLC "ยา 137" AT %MW1122, 1 s
   "ยา 138" : Word = PLC "ยา 138" AT %MW1124, 1 s
   "ยา 139" : Word = PLC "ยา 139" AT %MW1126, 1 s
   "ยา 14" : Word = PLC "ยา 14" AT %MW876, 1 s
   "ยา 140" : Word = PLC "ยา 140" AT %MW1128, 1 s
   "ยา 141" : Word = PLC "ยา 141" AT %MW1130, 1 s
   "ยา 142" : Word = PLC "ยา 142" AT %MW1132, 1 s
   "ยา 143" : Word = PLC "ยา 143" AT %MW1134, 1 s
   "ยา 144" : Word = PLC "ยา 144" AT %MW1136, 1 s
   "ยา 145" : Word = PLC "ยา 145" AT %MW1138, 1 s
   "ยา 146" : Word = PLC "ยา 146" AT %MW1140, 1 s
   "ยา 147" : Word = PLC "ยา 147" AT %MW1142, 1 s
   "ยา 148" : Word = PLC "ยา 148" AT %MW1144, 1 s
   "ยา 149" : Word = PLC "ยา 149" AT %MW1146, 1 s
   "ยา 15" : Word = PLC "ยา 15" AT %MW878, 1 s
   "ยา 150" : Word = PLC "ยา 150" AT %MW1148, 1 s
   "ยา 151" : Word = PLC "ยา 151" AT %MW1150, 1 s
   "ยา 152" : Word = PLC "ยา 152" AT %MW1152, 1 s
   "ยา 153" : Word = PLC "ยา 153" AT %MW1154, 1 s
   "ยา 154" : Word = PLC "ยา 154" AT %MW1156, 1 s
   "ยา 155" : Word = PLC "ยา 155" AT %MW1158, 1 s
   "ยา 156" : Word = PLC "ยา 156" AT %MW1160, 1 s
   "ยา 157" : Word = PLC "ยา 157" AT %MW1162, 1 s
   "ยา 158" : Word = PLC "ยา 158" AT %MW1164, 1 s
   "ยา 159" : Word = PLC "ยา 159" AT %MW1166, 1 s
   "ยา 16" : Word = PLC "ยา 16" AT %MW880, 1 s
   "ยา 160" : Word = PLC "ยา 160" AT %MW1168, 1 s
   "ยา 161" : Word = PLC "ยา 161" AT %MW1170, 1 s
   "ยา 162" : Word = PLC "ยา 162" AT %MW1172, 1 s
   "ยา 163" : Word = PLC "ยา 163" AT %MW1174, 1 s
   "ยา 164" : Word = PLC "ยา 164" AT %MW1890, 1 s
   "ยา 165" : Word = PLC "ยา 165" AT %MW1178, 1 s
   "ยา 166" : Word = PLC "ยา 166" AT %MW1180, 1 s
   "ยา 167" : Word = PLC "ยา 167" AT %MW1182, 1 s
   "ยา 168" : Word = PLC "ยา 168" AT %MW1184, 1 s
   "ยา 169" : Word = PLC "ยา 169" AT %MW1186, 1 s
   "ยา 17" : Word = PLC "ยา 17" AT %MW882, 1 s
   "ยา 170" : Word = PLC "ยา 170" AT %MW1188, 1 s
   "ยา 171" : Word = PLC "ยา 171" AT %MW1190, 1 s
   "ยา 172" : Word = PLC "ยา 172" AT %MW1192, 1 s
   "ยา 173" : Word = PLC "ยา 173" AT %MW1194, 1 s
   "ยา 174" : Word = PLC "ยา 174" AT %MW1196, 1 s
   "ยา 175" : Word = PLC "ยา 175" AT %MW1198, 1 s
   "ยา 176" : Word = PLC "ยา 176" AT %MW1200, 1 s
   "ยา 177" : Word = PLC "ยา 177" AT %MW1202, 1 s
   "ยา 178" : Word = PLC "ยา 178" AT %MW1204, 1 s
   "ยา 179" : Word = PLC "ยา 179" AT %MW1206, 1 s
   "ยา 18" : Word = PLC "ยา 18" AT %MW884, 1 s
   "ยา 180" : Word = PLC "ยา 180" AT %MW1208, 1 s
   "ยา 181" : Word = PLC "ยา 181" AT %MW1210, 1 s
   "ยา 182" : Word = PLC "ยา 182" AT %MW1212, 1 s
   "ยา 183" : Word = PLC "ยา 183" AT %MW1214, 1 s
   "ยา 184" : Word = PLC "ยา 184" AT %MW1216, 1 s
   "ยา 185" : Word = PLC "ยา 185" AT %MW1218, 1 s
   "ยา 186" : Word = PLC "ยา 186" AT %MW1220, 1 s
   "ยา 187" : Word = PLC "ยา 187" AT %MW1222, 1 s
   "ยา 188" : Word = PLC "ยา 188" AT %MW1224, 1 s
   "ยา 189" : Word = PLC "ยา 189" AT %MW1226, 1 s
   "ยา 19" : Word = PLC "ยา 19" AT %MW886, 1 s
   "ยา 190" : Word = PLC "ยา 190" AT %MW1228, 1 s
   "ยา 191" : Word = PLC "ยา 191" AT %MW1230, 1 s
   "ยา 192" : Word = PLC "ยา 192" AT %MW1232, 1 s
   "ยา 193" : Word = PLC "ยา 193" AT %MW1234, 1 s
   "ยา 194" : Word = PLC "ยา 194" AT %MW1236, 1 s
   "ยา 195" : Word = PLC "ยา 195" AT %MW1238, 1 s
   "ยา 196" : Word = PLC "ยา 196" AT %MW1240, 1 s
   "ยา 197" : Word = PLC "ยา 197" AT %MW1242, 1 s
   "ยา 198" : Word = PLC "ยา 198" AT %MW1244, 1 s
   "ยา 199" : Word = PLC "ยา 199" AT %MW1246, 1 s
   "ยา 2" : Word = PLC "ยา 2" AT %MW852, 1 s
   "ยา 20" : Word = PLC "ยา 20" AT %MW888, 1 s
   "ยา 200" : Word = PLC "ยา 200" AT %MW1248, 1 s
   "ยา 201" : Word = PLC "ยา 201" AT %MW1250, 1 s
   "ยา 202" : Word = PLC "ยา 202" AT %MW1252, 1 s
   "ยา 203" : Word = PLC "ยา 203" AT %MW1254, 1 s
   "ยา 204" : Word = PLC "ยา 204" AT %MW1256, 1 s
   "ยา 205" : Word = PLC "ยา 205" AT %MW1258, 1 s
   "ยา 206" : Word = PLC "ยา 206" AT %MW1260, 1 s
   "ยา 207" : Word = PLC "ยา 207" AT %MW1262, 1 s
   "ยา 208" : Word = PLC "ยา 208" AT %MW1264, 1 s
   "ยา 209" : Word = PLC "ยา 209" AT %MW1266, 1 s
   "ยา 21" : Word = PLC "ยา 21" AT %MW890, 1 s
   "ยา 210" : Word = PLC "ยา 210" AT %MW1268, 1 s
   "ยา 211" : Word = PLC "ยา 211" AT %MW1270, 1 s
   "ยา 212" : Word = PLC "ยา 212" AT %MW1272, 1 s
   "ยา 213" : Word = PLC "ยา 213" AT %MW1274, 1 s
   "ยา 214" : Word = PLC "ยา 214" AT %MW1276, 1 s
   "ยา 215" : Word = PLC "ยา 215" AT %MW1278, 1 s
   "ยา 216" : Word = PLC "ยา 216" AT %MW1280, 1 s
   "ยา 217" : Word = PLC "ยา 217" AT %MW1282, 1 s
   "ยา 218" : Word = PLC "ยา 218" AT %MW1284, 1 s
   "ยา 219" : Word = PLC "ยา 219" AT %MW1286, 1 s
   "ยา 22" : Word = PLC "ยา 22" AT %MW892, 1 s
   "ยา 220" : Word = PLC "ยา 220" AT %MW1288, 1 s
   "ยา 221" : Word = PLC "ยา 221" AT %MW1290, 1 s
   "ยา 222" : Word = PLC "ยา 222" AT %MW1292, 1 s
   "ยา 223" : Word = PLC "ยา 223" AT %MW1294, 1 s
   "ยา 224" : Word = PLC "ยา 224" AT %MW1296, 1 s
   "ยา 225" : Word = PLC "ยา 225" AT %MW1298, 1 s
   "ยา 226" : Word = PLC "ยา 226" AT %MW1300, 1 s
   "ยา 227" : Word = PLC "ยา 227" AT %MW1302, 1 s
   "ยา 228" : Word = PLC "ยา 228" AT %MW1304, 1 s
   "ยา 229" : Word = PLC "ยา 229" AT %MW1306, 1 s
   "ยา 23" : Word = PLC "ยา 23" AT %MW894, 1 s
   "ยา 230" : Word = PLC "ยา 230" AT %MW1308, 1 s
   "ยา 231" : Word = PLC "ยา 231" AT %MW1310, 1 s
   "ยา 232" : Word = PLC "ยา 232" AT %MW1312, 1 s
   "ยา 233" : Word = PLC "ยา 233" AT %MW1314, 1 s
   "ยา 234" : Word = PLC "ยา 234" AT %MW1316, 1 s
   "ยา 235" : Word = PLC "ยา 235" AT %MW1318, 1 s
   "ยา 236" : Word = PLC "ยา 236" AT %MW1320, 1 s
   "ยา 237" : Word = PLC "ยา 237" AT %MW1322, 1 s
   "ยา 238" : Word = PLC "ยา 238" AT %MW1324, 1 s
   "ยา 239" : Word = PLC "ยา 239" AT %MW1326, 1 s
   "ยา 24" : Word = PLC "ยา 24" AT %MW896, 1 s
   "ยา 240" : Word = PLC "ยา 240" AT %MW1328, 1 s
   "ยา 241" : Word = PLC "ยา 241" AT %MW1330, 1 s
   "ยา 242" : Word = PLC "ยา 242" AT %MW1332, 1 s
   "ยา 243" : Word = PLC "ยา 243" AT %MW1334, 1 s
   "ยา 244" : Word = PLC "ยา 244" AT %MW1336, 1 s
   "ยา 245" : Word = PLC "ยา 245" AT %MW1338, 1 s
   "ยา 246" : Word = PLC "ยา 246" AT %MW1340, 1 s
   "ยา 247" : Word = PLC "ยา 247" AT %MW1342, 1 s
   "ยา 248" : Word = PLC "ยา 248" AT %MW1344, 1 s
   "ยา 249" : Word = PLC "ยา 249" AT %MW1346, 1 s
   "ยา 25" : Word = PLC "ยา 25" AT %MW898, 1 s
   "ยา 250" : Word = PLC "ยา 250" AT %MW1348, 1 s
   "ยา 251" : Word = PLC "ยา 251" AT %MW1350, 1 s
   "ยา 252" : Word = PLC "ยา 252" AT %MW1352, 1 s
   "ยา 253" : Word = PLC "ยา 253" AT %MW1354, 1 s
   "ยา 254" : Word = PLC "ยา 254" AT %MW1356, 1 s
   "ยา 255" : Word = PLC "ยา 255" AT %MW1358, 1 s
   "ยา 256" : Word = PLC "ยา 256" AT %MW1360, 1 s
   "ยา 257" : Word = PLC "ยา 257" AT %MW1362, 1 s
   "ยา 258" : Word = PLC "ยา 258" AT %MW1364, 1 s
   "ยา 259" : Word = PLC "ยา 259" AT %MW1366, 1 s
   "ยา 26" : Word = PLC "ยา 26" AT %MW900, 1 s
   "ยา 260" : Word = PLC "ยา 260" AT %MW1368, 1 s
   "ยา 261" : Word = PLC "ยา 261" AT %MW1370, 1 s
   "ยา 262" : Word = PLC "ยา 262" AT %MW1372, 1 s
   "ยา 263" : Word = PLC "ยา 263" AT %MW1374, 1 s
   "ยา 264" : Word = PLC "ยา 264" AT %MW1376, 1 s
   "ยา 265" : Word = PLC "ยา 265" AT %MW1378, 1 s
   "ยา 266" : Word = PLC "ยา 266" AT %MW1380, 1 s
   "ยา 267" : Word = PLC "ยา 267" AT %MW1382, 1 s
   "ยา 268" : Word = PLC "ยา 268" AT %MW1384, 1 s
   "ยา 269" : Word = PLC "ยา 269" AT %MW1386, 1 s
   "ยา 27" : Word = PLC "ยา 27" AT %MW902, 1 s
   "ยา 270" : Word = PLC "ยา 270" AT %MW1388, 1 s
   "ยา 271" : Word = PLC "ยา 271" AT %MW1390, 1 s
   "ยา 272" : Word = PLC "ยา 272" AT %MW1392, 1 s
   "ยา 273" : Word = PLC "ยา 273" AT %MW1394, 1 s
   "ยา 274" : Word = PLC "ยา 274" AT %MW1396, 1 s
   "ยา 275" : Word = PLC "ยา 275" AT %MW1398, 1 s
   "ยา 276" : Word = PLC "ยา 276" AT %MW1400, 1 s
   "ยา 277" : Word = PLC "ยา 277" AT %MW1402, 1 s
   "ยา 278" : Word = PLC "ยา 278" AT %MW1404, 1 s
   "ยา 279" : Word = PLC "ยา 279" AT %MW1406, 1 s
   "ยา 28" : Word = PLC "ยา 28" AT %MW904, 1 s
   "ยา 280" : Word = PLC "ยา 280" AT %MW1408, 1 s
   "ยา 281" : Word = PLC "ยา 281" AT %MW1410, 1 s
   "ยา 282" : Word = PLC "ยา 282" AT %MW1412, 1 s
   "ยา 283" : Word = PLC "ยา 283" AT %MW1414, 1 s
   "ยา 284" : Word = PLC "ยา 284" AT %MW1416, 1 s
   "ยา 285" : Word = PLC "ยา 285" AT %MW1418, 1 s
   "ยา 286" : Word = PLC "ยา 286" AT %MW1420, 1 s
   "ยา 287" : Word = PLC "ยา 287" AT %MW1422, 1 s
   "ยา 288" : Word = PLC "ยา 288" AT %MW1424, 1 s
   "ยา 289" : Word = PLC "ยา 289" AT %MW1426, 1 s
   "ยา 29" : Word = PLC "ยา 29" AT %MW906, 1 s
   "ยา 290" : Word = PLC "ยา 290" AT %MW1428, 1 s
   "ยา 291" : Word = PLC "ยา 291" AT %MW1430, 1 s
   "ยา 292" : Word = PLC "ยา 292" AT %MW1432, 1 s
   "ยา 293" : Word = PLC "ยา 293" AT %MW1434, 1 s
   "ยา 294" : Word = PLC "ยา 294" AT %MW1436, 1 s
   "ยา 295" : Word = PLC "ยา 295" AT %MW1438, 1 s
   "ยา 296" : Word = PLC "ยา 296" AT %MW1440, 1 s
   "ยา 297" : Word = PLC "ยา 297" AT %MW1442, 1 s
   "ยา 298" : Word = PLC "ยา 298" AT %MW1444, 1 s
   "ยา 299" : Word = PLC "ยา 299" AT %MW1446, 1 s
   "ยา 3" : Word = PLC "ยา 3" AT %MW854, 1 s
   "ยา 30" : Word = PLC "ยา 30" AT %MW908, 1 s
   "ยา 300" : Word = PLC "ยา 300" AT %MW1448, 1 s
   "ยา 301" : Word = PLC "ยา 301" AT %MW1450, 1 s
   "ยา 302" : Word = PLC "ยา 302" AT %MW1452, 1 s
   "ยา 303" : Word = PLC "ยา 303" AT %MW1454, 1 s
   "ยา 304" : Word = PLC "ยา 304" AT %MW1456, 1 s
   "ยา 305" : Word = PLC "ยา 305" AT %MW1458, 1 s
   "ยา 306" : Word = PLC "ยา 306" AT %MW1460, 1 s
   "ยา 307" : Word = PLC "ยา 307" AT %MW1462, 1 s
   "ยา 308" : Word = PLC "ยา 308" AT %MW1464, 1 s
   "ยา 309" : Word = PLC "ยา 309" AT %MW1466, 1 s
   "ยา 31" : Word = PLC "ยา 31" AT %MW910, 1 s
   "ยา 310" : Word = PLC "ยา 310" AT %MW1468, 1 s
   "ยา 311" : Word = PLC "ยา 311" AT %MW1470, 1 s
   "ยา 312" : Word = PLC "ยา 312" AT %MW1472, 1 s
   "ยา 313" : Word = PLC "ยา 313" AT %MW1474, 1 s
   "ยา 314" : Word = PLC "ยา 314" AT %MW1476, 1 s
   "ยา 315" : Word = PLC "ยา 315" AT %MW1478, 1 s
   "ยา 316" : Word = PLC "ยา 316" AT %MW1480, 1 s
   "ยา 317" : Word = PLC "ยา 317" AT %MW1482, 1 s
   "ยา 318" : Word = PLC "ยา 318" AT %MW1484, 1 s
   "ยา 319" : Word = PLC "ยา 319" AT %MW1486, 1 s
   "ยา 32" : Word = PLC "ยา 32" AT %MW912, 1 s
   "ยา 320" : Word = PLC "ยา 320" AT %MW1488, 1 s
   "ยา 321" : Word = PLC "ยา 321" AT %MW1490, 1 s
   "ยา 322" : Word = PLC "ยา 322" AT %MW1492, 1 s
   "ยา 323" : Word = PLC "ยา 323" AT %MW1494, 1 s
   "ยา 324" : Word = PLC "ยา 324" AT %MW1496, 1 s
   "ยา 325" : Word = PLC "ยา 325" AT %MW1498, 1 s
   "ยา 326" : Word = PLC "ยา 326" AT %MW1500, 1 s
   "ยา 327" : Word = PLC "ยา 327" AT %MW1502, 1 s
   "ยา 328" : Word = PLC "ยา 328" AT %MW1504, 1 s
   "ยา 329" : Word = PLC "ยา 329" AT %MW1506, 1 s
   "ยา 33" : Word = PLC "ยา 33" AT %MW914, 1 s
   "ยา 330" : Word = PLC "ยา 330" AT %MW1508, 1 s
   "ยา 331" : Word = PLC "ยา 331" AT %MW1510, 1 s
   "ยา 332" : Word = PLC "ยา 332" AT %MW1512, 1 s
   "ยา 333" : Word = PLC "ยา 333" AT %MW1514, 1 s
   "ยา 334" : Word = PLC "ยา 334" AT %MW1516, 1 s
   "ยา 335" : Word = PLC "ยา 335" AT %MW1518, 1 s
   "ยา 336" : Word = PLC "ยา 336" AT %MW1520, 1 s
   "ยา 337" : Word = PLC "ยา 337" AT %MW1522, 1 s
   "ยา 338" : Word = PLC "ยา 338" AT %MW1524, 1 s
   "ยา 339" : Word = PLC "ยา 339" AT %MW1526, 1 s
   "ยา 34" : Word = PLC "ยา 34" AT %MW916, 1 s
   "ยา 340" : Word = PLC "ยา 340" AT %MW1528, 1 s
   "ยา 341" : Word = PLC "ยา 341" AT %MW1530, 1 s
   "ยา 342" : Word = PLC "ยา 342" AT %MW1532, 1 s
   "ยา 343" : Word = PLC "ยา 343" AT %MW1534, 1 s
   "ยา 344" : Word = PLC "ยา 344" AT %MW1536, 1 s
   "ยา 345" : Word = PLC "ยา 345" AT %MW1538, 1 s
   "ยา 346" : Word = PLC "ยา 346" AT %MW1540, 1 s
   "ยา 347" : Word = PLC "ยา 347" AT %MW1542, 1 s
   "ยา 348" : Word = PLC "ยา 348" AT %MW1544, 1 s
   "ยา 349" : Word = PLC "ยา 349" AT %MW1546, 1 s
   "ยา 35" : Word = PLC "ยา 35" AT %MW918, 1 s
   "ยา 350" : Word = PLC "ยา 350" AT %MW1548, 1 s
   "ยา 351" : Word = PLC "ยา 351" AT %MW1550, 1 s
   "ยา 352" : Word = PLC "ยา 352" AT %MW1552, 1 s
   "ยา 353" : Word = PLC "ยา 353" AT %MW1554, 1 s
   "ยา 354" : Word = PLC "ยา 354" AT %MW1556, 1 s
   "ยา 355" : Word = PLC "ยา 355" AT %MW1558, 1 s
   "ยา 356" : Word = PLC "ยา 356" AT %MW1560, 1 s
   "ยา 357" : Word = PLC "ยา 357" AT %MW1562, 1 s
   "ยา 358" : Word = PLC "ยา 358" AT %MW1564, 1 s
   "ยา 359" : Word = PLC "ยา 359" AT %MW1566, 1 s
   "ยา 36" : Word = PLC "ยา 36" AT %MW920, 1 s
   "ยา 360" : Word = PLC "ยา 360" AT %MW1568, 1 s
   "ยา 361" : Word = PLC "ยา 361" AT %MW1570, 1 s
   "ยา 362" : Word = PLC "ยา 362" AT %MW1572, 1 s
   "ยา 363" : Word = PLC "ยา 363" AT %MW1574, 1 s
   "ยา 364" : Word = PLC "ยา 364" AT %MW1576, 1 s
   "ยา 365" : Word = PLC "ยา 365" AT %MW1578, 1 s
   "ยา 366" : Word = PLC "ยา 366" AT %MW1580, 1 s
   "ยา 367" : Word = PLC "ยา 367" AT %MW1582, 1 s
   "ยา 368" : Word = PLC "ยา 368" AT %MW1584, 1 s
   "ยา 369" : Word = PLC "ยา 369" AT %MW1586, 1 s
   "ยา 37" : Word = PLC "ยา 37" AT %MW922, 1 s
   "ยา 370" : Word = PLC "ยา 370" AT %MW1588, 1 s
   "ยา 371" : Word = PLC "ยา 371" AT %MW1590, 1 s
   "ยา 372" : Word = PLC "ยา 372" AT %MW1592, 1 s
   "ยา 373" : Word = PLC "ยา 373" AT %MW1594, 1 s
   "ยา 374" : Word = PLC "ยา 374" AT %MW1596, 1 s
   "ยา 375" : Word = PLC "ยา 375" AT %MW1598, 1 s
   "ยา 376" : Word = PLC "ยา 376" AT %MW1600, 1 s
   "ยา 377" : Word = PLC "ยา 377" AT %MW1602, 1 s
   "ยา 378" : Word = PLC "ยา 378" AT %MW1604, 1 s
   "ยา 379" : Word = PLC "ยา 379" AT %MW1606, 1 s
   "ยา 38" : Word = PLC "ยา 38" AT %MW924, 1 s
   "ยา 380" : Word = PLC "ยา 380" AT %MW1608, 1 s
   "ยา 381" : Word = PLC "ยา 381" AT %MW1610, 1 s
   "ยา 382" : Word = PLC "ยา 382" AT %MW1612, 1 s
   "ยา 383" : Word = PLC "ยา 383" AT %MW1614, 1 s
   "ยา 384" : Word = PLC "ยา 384" AT %MW1616, 1 s
   "ยา 385" : Word = PLC "ยา 385" AT %MW1618, 1 s
   "ยา 386" : Word = PLC "ยา 386" AT %MW1620, 1 s
   "ยา 387" : Word = PLC "ยา 387" AT %MW1622, 1 s
   "ยา 388" : Word = PLC "ยา 388" AT %MW1624, 1 s
   "ยา 389" : Word = PLC "ยา 389" AT %MW1626, 1 s
   "ยา 39" : Word = PLC "ยา 39" AT %MW926, 1 s
   "ยา 390" : Word = PLC "ยา 390" AT %MW1628, 1 s
   "ยา 391" : Word = PLC "ยา 391" AT %MW1630, 1 s
   "ยา 392" : Word = PLC "ยา 392" AT %MW1632, 1 s
   "ยา 393" : Word = PLC "ยา 393" AT %MW1634, 1 s
   "ยา 394" : Word = PLC "ยา 394" AT %MW1636, 1 s
   "ยา 395" : Word = PLC "ยา 395" AT %MW1638, 1 s
   "ยา 396" : Word = PLC "ยา 396" AT %MW1640, 1 s
   "ยา 397" : Word = PLC "ยา 397" AT %MW1642, 1 s
   "ยา 398" : Word = PLC "ยา 398" AT %MW1644, 1 s
   "ยา 399" : Word = PLC "ยา 399" AT %MW1646, 1 s
   "ยา 4" : Word = PLC "ยา 4" AT %MW856, 1 s
   "ยา 40" : Word = PLC "ยา 40" AT %MW928, 1 s
   "ยา 400" : Word = PLC "ยา 400" AT %MW1648, 1 s
   "ยา 401" : Word = PLC "ยา 401" AT %MW1650, 1 s
   "ยา 402" : Word = PLC "ยา 402" AT %MW1652, 1 s
   "ยา 403" : Word = PLC "ยา 403" AT %MW1654, 1 s
   "ยา 404" : Word = PLC "ยา 404" AT %MW1656, 1 s
   "ยา 405" : Word = PLC "ยา 405" AT %MW1658, 1 s
   "ยา 406" : Word = PLC "ยา 406" AT %MW1660, 1 s
   "ยา 407" : Word = PLC "ยา 407" AT %MW1662, 1 s
   "ยา 408" : Word = PLC "ยา 408" AT %MW1664, 1 s
   "ยา 409" : Word = PLC "ยา 409" AT %MW1666, 1 s
   "ยา 41" : Word = PLC "ยา 41" AT %MW930, 1 s
   "ยา 410" : Word = PLC "ยา 410" AT %MW1668, 1 s
   "ยา 411" : Word = PLC "ยา 411" AT %MW1670, 1 s
   "ยา 412" : Word = PLC "ยา 412" AT %MW1672, 1 s
   "ยา 413" : Word = PLC "ยา 413" AT %MW1674, 1 s
   "ยา 414" : Word = PLC "ยา 414" AT %MW1676, 1 s
   "ยา 415" : Word = PLC "ยา 415" AT %MW1678, 1 s
   "ยา 416" : Word = PLC "ยา 416" AT %MW1680, 1 s
   "ยา 417" : Word = PLC "ยา 417" AT %MW1682, 1 s
   "ยา 418" : Word = PLC "ยา 418" AT %MW1684, 1 s
   "ยา 419" : Word = PLC "ยา 419" AT %MW1686, 1 s
   "ยา 42" : Word = PLC "ยา 42" AT %MW932, 1 s
   "ยา 420" : Word = PLC "ยา 420" AT %MW1688, 1 s
   "ยา 421" : Word = PLC "ยา 421" AT %MW1690, 1 s
   "ยา 422" : Word = PLC "ยา 422" AT %MW1692, 1 s
   "ยา 423" : Word = PLC "ยา 423" AT %MW1694, 1 s
   "ยา 424" : Word = PLC "ยา 424" AT %MW1696, 1 s
   "ยา 425" : Word = PLC "ยา 425" AT %MW1698, 1 s
   "ยา 426" : Word = PLC "ยา 426" AT %MW1700, 1 s
   "ยา 427" : Word = PLC "ยา 427" AT %MW1702, 1 s
   "ยา 428" : Word = PLC "ยา 428" AT %MW1704, 1 s
   "ยา 429" : Word = PLC "ยา 429" AT %MW1706, 1 s
   "ยา 43" : Word = PLC "ยา 43" AT %MW934, 1 s
   "ยา 430" : Word = PLC "ยา 430" AT %MW1708, 1 s
   "ยา 431" : Word = PLC "ยา 431" AT %MW1710, 1 s
   "ยา 432" : Word = PLC "ยา 432" AT %MW1712, 1 s
   "ยา 433" : Word = PLC "ยา 433" AT %MW1714, 1 s
   "ยา 434" : Word = PLC "ยา 434" AT %MW1716, 1 s
   "ยา 435" : Word = PLC "ยา 435" AT %MW1718, 1 s
   "ยา 436" : Word = PLC "ยา 436" AT %MW1720, 1 s
   "ยา 437" : Word = PLC "ยา 437" AT %MW1722, 1 s
   "ยา 438" : Word = PLC "ยา 438" AT %MW1724, 1 s
   "ยา 439" : Word = PLC "ยา 439" AT %MW1726, 1 s
   "ยา 44" : Word = PLC "ยา 44" AT %MW936, 1 s
   "ยา 440" : Word = PLC "ยา 440" AT %MW1728, 1 s
   "ยา 441" : Word = PLC "ยา 441" AT %MW1730, 1 s
   "ยา 442" : Word = PLC "ยา 442" AT %MW1732, 1 s
   "ยา 443" : Word = PLC "ยา 443" AT %MW1734, 1 s
   "ยา 444" : Word = PLC "ยา 444" AT %MW1736, 1 s
   "ยา 445" : Word = PLC "ยา 445" AT %MW1738, 1 s
   "ยา 446" : Word = PLC "ยา 446" AT %MW1740, 1 s
   "ยา 447" : Word = PLC "ยา 447" AT %MW1742, 1 s
   "ยา 448" : Word = PLC "ยา 448" AT %MW1744, 1 s
   "ยา 449" : Word = PLC "ยา 449" AT %MW1746, 1 s
   "ยา 45" : Word = PLC "ยา 45" AT %MW938, 1 s
   "ยา 450" : Word = PLC "ยา 450" AT %MW1748, 1 s
   "ยา 451" : Word = PLC "ยา 451" AT %MW1750, 1 s
   "ยา 452" : Word = PLC "ยา 452" AT %MW1752, 1 s
   "ยา 453" : Word = PLC "ยา 453" AT %MW1754, 1 s
   "ยา 454" : Word = PLC "ยา 454" AT %MW1756, 1 s
   "ยา 455" : Word = PLC "ยา 455" AT %MW1758, 1 s
   "ยา 456" : Word = PLC "ยา 456" AT %MW1760, 1 s
   "ยา 457" : Word = PLC "ยา 457" AT %MW1762, 1 s
   "ยา 458" : Word = PLC "ยา 458" AT %MW1764, 1 s
   "ยา 459" : Word = PLC "ยา 459" AT %MW1766, 1 s
   "ยา 46" : Word = PLC "ยา 46" AT %MW940, 1 s
   "ยา 460" : Word = PLC "ยา 460" AT %MW1768, 1 s
   "ยา 461" : Word = PLC "ยา 461" AT %MW1770, 1 s
   "ยา 462" : Word = PLC "ยา 462" AT %MW1772, 1 s
   "ยา 463" : Word = PLC "ยา 463" AT %MW1774, 1 s
   "ยา 464" : Word = PLC "ยา 464" AT %MW1776, 1 s
   "ยา 465" : Word = PLC "ยา 465" AT %MW1778, 1 s
   "ยา 466" : Word = PLC "ยา 466" AT %MW1780, 1 s
   "ยา 467" : Word = PLC "ยา 467" AT %MW1782, 1 s
   "ยา 468" : Word = PLC "ยา 468" AT %MW1784, 1 s
   "ยา 469" : Word = PLC "ยา 469" AT %MW1786, 1 s
   "ยา 47" : Word = PLC "ยา 47" AT %MW942, 1 s
   "ยา 470" : Word = PLC "ยา 470" AT %MW1788, 1 s
   "ยา 471" : Word = PLC "ยา 471" AT %MW1790, 1 s
   "ยา 472" : Word = PLC "ยา 472" AT %MW1792, 1 s
   "ยา 473" : Word = PLC "ยา 473" AT %MW1794, 1 s
   "ยา 474" : Word = PLC "ยา 474" AT %MW1796, 1 s
   "ยา 475" : Word = PLC "ยา 475" AT %MW1798, 1 s
   "ยา 476" : Word = PLC "ยา 476" AT %MW1800, 1 s
   "ยา 477" : Word = PLC "ยา 477" AT %MW1802, 1 s
   "ยา 478" : Word = PLC "ยา 478" AT %MW1804, 1 s
   "ยา 479" : Word = PLC "ยา 479" AT %MW1806, 1 s
   "ยา 48" : Word = PLC "ยา 48" AT %MW944, 1 s
   "ยา 480" : Word = PLC "ยา 480" AT %MW1808, 1 s
   "ยา 481" : Word = PLC "ยา 481" AT %MW1810, 1 s
   "ยา 482" : Word = PLC "ยา 482" AT %MW1812, 1 s
   "ยา 483" : Word = PLC "ยา 483" AT %MW1814, 1 s
   "ยา 484" : Word = PLC "ยา 484" AT %MW1816, 1 s
   "ยา 485" : Word = PLC "ยา 485" AT %MW1818, 1 s
   "ยา 486" : Word = PLC "ยา 486" AT %MW1820, 1 s
   "ยา 487" : Word = PLC "ยา 487" AT %MW1822, 1 s
   "ยา 488" : Word = PLC "ยา 488" AT %MW1824, 1 s
   "ยา 489" : Word = PLC "ยา 489" AT %MW1826, 1 s
   "ยา 49" : Word = PLC "ยา 49" AT %MW946, 1 s
   "ยา 490" : Word = PLC "ยา 490" AT %MW1828, 1 s
   "ยา 491" : Word = PLC "ยา 491" AT %MW1830, 1 s
   "ยา 492" : Word = PLC "ยา 492" AT %MW1832, 1 s
   "ยา 493" : Word = PLC "ยา 493" AT %MW1834, 1 s
   "ยา 494" : Word = PLC "ยา 494" AT %MW1836, 1 s
   "ยา 495" : Word = PLC "ยา 495" AT %MW1838, 1 s
   "ยา 496" : Word = PLC "ยา 496" AT %MW1840, 1 s
   "ยา 497" : Word = PLC "ยา 497" AT %MW1842, 1 s
   "ยา 498" : Word = PLC "ยา 498" AT %MW1844, 1 s
   "ยา 499" : Word = PLC "ยา 499" AT %MW1846, 1 s
   "ยา 5" : Word = PLC "ยา 5" AT %MW858, 1 s
   "ยา 50" : Word = PLC "ยา 50" AT %MW948, 1 s
   "ยา 500" : Word = PLC "ยา 500" AT %MW1848, 1 s
   "ยา 501" : Word = PLC "ยา 501" AT %MW1850, 1 s
   "ยา 502" : Word = PLC "ยา 502" AT %MW1852, 1 s
   "ยา 503" : Word = PLC "ยา 503" AT %MW1854, 1 s
   "ยา 504" : Word = PLC "ยา 504" AT %MW1856, 1 s
   "ยา 505" : Word = PLC "ยา 505" AT %MW1858, 1 s
   "ยา 506" : Word = PLC "ยา 506" AT %MW1860, 1 s
   "ยา 507" : Word = PLC "ยา 507" AT %MW1862, 1 s
   "ยา 508" : Word = PLC "ยา 508" AT %MW1864, 1 s
   "ยา 509" : Word = PLC "ยา 509" AT %MW1866, 1 s
   "ยา 51" : Word = PLC "ยา 51" AT %MW950, 1 s
   "ยา 510" : Word = PLC "ยา 510" AT %MW1868, 1 s
   "ยา 511" : Word = PLC "ยา 511" AT %MW1870, 1 s
   "ยา 512" : Word = PLC "ยา 512" AT %MW1872, 1 s
   "ยา 513" : Word = PLC "ยา 513" AT %MW1874, 1 s
   "ยา 514" : Word = PLC "ยา 514" AT %MW1876, 1 s
   "ยา 515" : Word = PLC "ยา 515" AT %MW1878, 1 s
   "ยา 516" : Word = PLC "ยา 516" AT %MW1880, 1 s
   "ยา 517" : Word = PLC "ยา 517" AT %MW1882, 1 s
   "ยา 518" : Word = PLC "ยา 518" AT %MW1884, 1 s
   "ยา 519" : Word = PLC "ยา 519" AT %MW1886, 1 s
   "ยา 52" : Word = PLC "ยา 52" AT %MW952, 1 s
   "ยา 520" : Word = PLC "ยา 520" AT %MW1888, 1 s
   "ยา 53" : Word = PLC "ยา 53" AT %MW954, 1 s
   "ยา 54" : Word = PLC "ยา 54" AT %MW956, 1 s
   "ยา 55" : Word = PLC "ยา 55" AT %MW958, 1 s
   "ยา 56" : Word = PLC "ยา 56" AT %MW960, 1 s
   "ยา 57" : Word = PLC "ยา 57" AT %MW962, 1 s
   "ยา 58" : Word = PLC "ยา 58" AT %MW964, 1 s
   "ยา 59" : Word = PLC "ยา 59" AT %MW966, 1 s
   "ยา 6" : Word = PLC "ยา 6" AT %MW860, 1 s
   "ยา 60" : Word = PLC "ยา 60" AT %MW968, 1 s
   "ยา 61" : Word = PLC "ยา 61" AT %MW970, 1 s
   "ยา 62" : Word = PLC "ยา 62" AT %MW972, 1 s
   "ยา 63" : Word = PLC "ยา 63" AT %MW974, 1 s
   "ยา 64" : Word = PLC "ยา 64" AT %MW976, 1 s
   "ยา 65" : Word = PLC "ยา 65" AT %MW978, 1 s
   "ยา 66" : Word = PLC "ยา 66" AT %MW980, 1 s
   "ยา 67" : Word = PLC "ยา 67" AT %MW982, 1 s
   "ยา 68" : Word = PLC "ยา 68" AT %MW984, 1 s
   "ยา 69" : Word = PLC "ยา 69" AT %MW986, 1 s
   "ยา 7" : Word = PLC "ยา 7" AT %MW862, 1 s
   "ยา 70" : Word = PLC "ยา 70" AT %MW988, 1 s
   "ยา 71" : Word = PLC "ยา 71" AT %MW990, 1 s
   "ยา 72" : Word = PLC "ยา 72" AT %MW992, 1 s
   "ยา 73" : Word = PLC "ยา 73" AT %MW994, 1 s
   "ยา 74" : Word = PLC "ยา 74" AT %MW996, 1 s
   "ยา 75" : Word = PLC "ยา 75" AT %MW998, 1 s
   "ยา 76" : Word = PLC "ยา 76" AT %MW1000, 1 s
   "ยา 77" : Word = PLC "ยา 77" AT %MW1002, 1 s
   "ยา 78" : Word = PLC "ยา 78" AT %MW1004, 1 s
   "ยา 79" : Word = PLC "ยา 79" AT %MW1006, 1 s
   "ยา 8" : Word = PLC "ยา 8" AT %MW864, 1 s
   "ยา 80" : Word = PLC "ยา 80" AT %MW1008, 1 s
   "ยา 81" : Word = PLC "ยา 81" AT %MW1010, 1 s
   "ยา 82" : Word = PLC "ยา 82" AT %MW1012, 1 s
   "ยา 83" : Word = PLC "ยา 83" AT %MW1014, 1 s
   "ยา 84" : Word = PLC "ยา 84" AT %MW1016, 1 s
   "ยา 85" : Word = PLC "ยา 85" AT %MW1018, 1 s
   "ยา 86" : Word = PLC "ยา 86" AT %MW1020, 1 s
   "ยา 87" : Word = PLC "ยา 87" AT %MW1022, 1 s
   "ยา 88" : Word = PLC "ยา 88" AT %MW1024, 1 s
   "ยา 89" : Word = PLC "ยา 89" AT %MW1026, 1 s
   "ยา 9" : Word = PLC "ยา 9" AT %MW866, 1 s
   "ยา 90" : Word = PLC "ยา 90" AT %MW1028, 1 s
   "ยา 91" : Word = PLC "ยา 91" AT %MW1030, 1 s
   "ยา 92" : Word = PLC "ยา 92" AT %MW1032, 1 s
   "ยา 93" : Word = PLC "ยา 93" AT %MW1034, 1 s
   "ยา 94" : Word = PLC "ยา 94" AT %MW1036, 1 s
   "ยา 95" : Word = PLC "ยา 95" AT %MW1038, 1 s
   "ยา 96" : Word = PLC "ยา 96" AT %MW1040, 1 s
   "ยา 97" : Word = PLC "ยา 97" AT %MW1042, 1 s
   "ยา 98" : Word = PLC "ยา 98" AT %MW1044, 1 s
   "ยา 99" : Word = PLC "ยา 99" AT %MW1046, 1 s
   "รอคำสั่งเบิกยา" : Bool = PLC รอคำสั่งเบิกยา AT %I102.0, 1 s
   "รอรับคำสั่งยา" : Bool = PLC รอรับคำสั่งยา AT %I101.3, 1 s
   "รับคำสั่งเบิกยา" : Bool = PLC รับคำสั่งเบิกยา AT %I101.4, 1 s
   "Emergency stop" : Bool = PLC "Emergency stop" AT %M1898.5, 1 s
   "Reset-All System" : Bool = PLC "Reset-All System" AT %M1898.6, 1 s

discrete alarms
   1: 'คอนเวเยอร์ Brushless Motor_NO', class Errors, trigger "Alarms_All" bit 0
   2: 'Stepper Motor ( PKP243D15A2-R2EL ) No.1_NO จัดเก็บ', class Errors, trigger "Alarms_All" bit 1
   3: 'Stepper Motor ( PKP243D15A2-R2EL )No.2_NO จัดเก็บ', class Errors, trigger "Alarms_All" bit 2
   4: 'Stepper motor + Gearhead ( PKP243D15A2-R2EL + PLE40-10B )_NO.3 จัดเก็บ', class Errors, trigger "Alarms_All" bit 3
   5: 'Stepper motor ( leadshine Nema24 CS-M22430) No.1_No จัดเก็บ', class Errors, trigger "Alarms_All" bit 4
   6: 'Stepper motor ( leadshine Nema24 CS-M22430) No.2_No จัดเก็บ', class Errors, trigger "Alarms_All" bit 5
   7: 'Stepper motor ( leadshine Nema24 CS-M22430) No.3_No จัดเก็บ', class Errors, trigger "Alarms_All" bit 6
   8: 'Stepper motor ( leadshine Nema24 CS-M22430) No.1 เบิกจ่าย', class Errors, trigger "Alarms_All" bit 7
   9: 'Stepper motor ( leadshine Nema24 CS-M22430) No.2 เบิกจ่าย', class Errors, trigger "Alarms_All" bit 8
   10: 'Stepper motor ( leadshine Nema24 CS-M22430) No.3 เบิกจ่าย', class Errors, trigger "Alarms_All" bit 9
   11: 'Stepper motor + Gearhead ( บริเวณกริปเปอร์ เบิกจ่าย )_No', class Errors, trigger "Alarms_All" bit 10
   12: 'Stepper motor ( บริเวณ คอนเวเยอร์ เบิกจ่าย )_No', class Errors, trigger "Alarms_All" bit 11
   13: 'Photoelectic sensor 1_จัดเก็บ_No', class Errors, trigger "Alarms_All" bit 12
   14: 'Photoelectic sensor 2_จัดเก็บ_No', class Errors, trigger "Alarms_All" bit 13
   15: 'Photoelectic Sensor No.1 เบิกจ่าย_No', class Errors, trigger "Alarms_All" bit 14
   16: 'Photoelectic Sensor No.2 เบิกจ่าย_No', class Errors, trigger "Alarms_All" bit 15

text list "Zone_y1.6": 0 'F'; 1 'L'; 2 'R'; 3 'X'

text list "Zone_y1.2": 0 'B'; 1 'H'; 2 'N'; 3 'T'; 4 'Z'

text list "Zone_y1.1": 0 'A'; 1 'G'; 2 'M'; 3 'S'; 4 'Y'

text list "Zone_x 1.3": 0 '3'; 1 '10'; 2 '17'

text list "Zone_y1.4": 0 'D'; 1 'J'; 2 'P'; 3 'V'

text list "Zone_x 1.7": 0 '7'; 1 '14'

text list "Zone_x 1.4": 0 '4'; 1 '11'; 2 '18'

text list "Zone_x 1.5": 0 '5'; 1 '12'; 2 '19'

text list "Zone_y1.3": 0 'C'; 1 'I'; 2 'O'; 3 'U'

text list "Zone_x 1.6": 0 '6'; 1 '13'; 2 '20'

text list "Zone_x 1.2": 0 '2'; 1 '9'; 2 '16'

text list "BOX_All": 1 'Box_1'; 2 'Box_2'; 3 'Box_3'; 4 'Box_4'; 5 'Box_5'; 6 'Box_6'; 7 'Box_7'; 8 'Box_8'; 9 'Box_9'; 10 'Box_10'; 11 'Box_11'; 12 'Box_12'; 13 'Box_13'; 14 'Box_14'; 15 'Box_15'; 16 'Box_16'; 17 'Box_17'; 18 'Box_18'; 19 'Box_19'; 20 'Box_20'; 21 'Box_21'; 22 'Box_22'; 23 'Box_23'; 24 'Box_24'; 25 'Box_25'; 26 'Box_26'; 27 'Box_27'; 28 'Box_28'; 29 'Box_29'; 30 'Box_30'; 31 'Box_31'; 32 'Box_32'; 33 'Box_33'; 34 'Box_34'; 35 'Box_35'; 36 'Box_36'; 37 'Box_37'; 38 'Box_38'; 39 'Box_39'; 40 'Box_40'; 41 'Box_41'; 42 'Box_42'; 43 'Box_43'; 44 'Box_44'; 45 'Box_45'; 46 'Box_46'; 47 'Box_47'; 48 'Box_48'; 49 'Box_49'; 50 'Box_50'; 51 'Box_51'; 52 'Box_52'; 53 'Box_53'; 54 'Box_54'; 55 'Box_55'; 56 'Box_56'; 57 'Box_57'; 58 'Box_58'; 59 'Box_59'; 60 'Box_60'; 61 'Box_61'; 62 'Box_62'; 63 'Box_63'; 64 'Box_64'; 65 'Box_65'; 66 'Box_66'; 67 'Box_67'; 68 'Box_68'; 69 'Box_69'; 70 'Box_70'; 71 'Box_71'; 72 'Box_72'; 73 'Box_73'; 74 'Box_74'; 75 'Box_75'; 76 'Box_76'; 77 'Box_77'; 78 'Box_78'; 79 'Box_79'; 80 'Box_80'; 81 'Box_81'; 82 'Box_82'; 83 'Box_83'; 84 'Box_84'; 85 'Box_85'; 86 'Box_86'; 87 'Box_87'; 88 'Box_88'; 89 'Box_89'; 90 'Box_90'; 91 'Box_91'; 92 'Box_92'; 93 'Box_93'; 94 'Box_94'; 95 'Box_95'; 96 'Box_96'; 97 'Box_97'; 98 'Box_98'; 99 'Box_99'; 100 'Box_100'; 101 'Box_101'; 102 'Box_102'; 103 'Box_103'; 104 'Box_104'; 105 'Box_105'; 106 'Box_106'; 107 'Box_107'; 108 'Box_108'; 109 'Box_109'; 110 'Box_110'; 111 'Box_111'; 112 'Box_112'; 113 'Box_113'; 114 'Box_114'; 115 'Box_115'; 116 'Box_116'; 117 'Box_117'; 118 'Box_118'; 119 'Box_119'; 120 'Box_120'; 121 'Box_121'; 122 'Box_122'; 123 'Box_123'; 124 'Box_124'; 125 'Box_125'; 126 'Box_126'; 127 'Box_127'; 128 'Box_128'; 129 'Box_129'; 130 'Box_130'; 131 'Box_131'; 132 'Box_132'; 133 'Box_133'; 134 'Box_134'; 135 'Box_135'; 136 'Box_136'; 137 'Box_137'; 138 'Box_138'; 139 'Box_139'; 140 'Box_140'; 141 'Box_141'; 142 'Box_142'; 143 'Box_143'; 144 'Box_144'; 145 'Box_145'; 146 'Box_146'; 147 'Box_147'; 148 'Box_148'; 149 'Box_149'; 150 'Box_150'; 151 'Box_151'; 152 'Box_152'; 153 'Box_153'; 154 'Box_154'; 155 'Box_155'; 156 'Box_156'; 157 'Box_157'; 158 'Box_158'; 159 'Box_159'; 160 'Box_160'; 161 'Box_161'; 162 'Box_162'; 163 'Box_163'; 164 'Box_164'; 165 'Box_165'; 166 'Box_166'; 167 'Box_167'; 168 'Box_168'; 169 'Box_169'; 170 'Box_170'; 171 'Box_171'; 172 'Box_172'; 173 'Box_173'; 174 'Box_174'; 175 'Box_175'; 176 'Box_176'; 177 'Box_177'; 178 'Box_178'; 179 'Box_179'; 180 'Box_180'; 181 'Box_181'; 182 'Box_182'; 183 'Box_183'; 184 'Box_184'; 185 'Box_185'; 186 'Box_186'; 187 'Box_187'; 188 'Box_188'; 189 'Box_189'; 190 'Box_190'; 191 'Box_191'; 192 'Box_192'; 193 'Box_193'; 194 'Box_194'; 195 'Box_195'; 196 'Box_196'; 197 'Box_197'; 198 'Box_198'; 199 'Box_199'; 200 'Box_200'; 201 'Box_201'; 202 'Box_202'; 203 'Box_203'; 204 'Box_204'; 205 'Box_205'; 206 'Box_206'; 207 'Box_207'; 208 'Box_208'; 209 'Box_209'; 210 'Box_210'; 211 'Box_211'; 212 'Box_212'; 213 'Box_213'; 214 'Box_214'; 215 'Box_215'; 216 'Box_216'; 217 'Box_217'; 218 'Box_218'; 219 'Box_219'; 220 'Box_220'; 221 'Box_221'; 222 'Box_222'; 223 'Box_223'; 224 'Box_224'; 225 'Box_225'; 226 'Box_226'; 227 'Box_227'; 228 'Box_228'; 229 'Box_229'; 230 'Box_230'; 231 'Box_231'; 232 'Box_232'; 233 'Box_233'; 234 'Box_234'; 235 'Box_235'; 236 'Box_236'; 237 'Box_237'; 238 'Box_238'; 239 'Box_239'; 240 'Box_240'; 241 'Box_241'; 242 'Box_242'; 243 'Box_243'; 244 'Box_244'; 245 'Box_245'; 246 'Box_246'; 247 'Box_247'; 248 'Box_248'; 249 'Box_249'; 250 'Box_250'; 251 'Box_251'; 252 'Box_252'; 253 'Box_253'; 254 'Box_254'; 255 'Box_255'; 256 'Box_256'; 257 'Box_257'; 258 'Box_258'; 259 'Box_259'; 260 'Box_260'; 261 'Box_261'; 262 'Box_262'; 263 'Box_263'; 264 'Box_264'; 265 'Box_265'; 266 'Box_266'; 267 'Box_267'; 268 'Box_268'; 269 'Box_269'; 270 'Box_270'; 271 'Box_271'; 272 'Box_272'; 273 'Box_273'; 274 'Box_274'; 275 'Box_275'; 276 'Box_276'; 277 'Box_277'; 278 'Box_278'; 279 'Box_279'; 280 'Box_280'; 281 'Box_281'; 282 'Box_282'; 283 'Box_283'; 284 'Box_284'; 285 'Box_285'; 286 'Box_286'; 287 'Box_287'; 288 'Box_288'; 289 'Box_289'; 290 'Box_290'; 291 'Box_291'; 292 'Box_292'; 293 'Box_293'; 294 'Box_294'; 295 'Box_295'; 296 'Box_296'; 297 'Box_297'; 298 'Box_298'; 299 'Box_299'; 300 'Box_300'; 301 'Box_301'; 302 'Box_302'; 303 'Box_303'; 304 'Box_304'; 305 'Box_305'; 306 'Box_306'; 307 'Box_307'; 308 'Box_308'; 309 'Box_309'; 310 'Box_310'; 311 'Box_311'; 312 'Box_312'; 313 'Box_313'; 314 'Box_314'; 315 'Box_315'; 316 'Box_316'; 317 'Box_317'; 318 'Box_318'; 319 'Box_319'; 320 'Box_320'; 321 'Box_321'; 322 'Box_322'; 323 'Box_323'; 324 'Box_324'; 325 'Box_325'; 326 'Box_326'; 327 'Box_327'; 328 'Box_328'; 329 'Box_329'; 330 'Box_330'; 331 'Box_331'; 332 'Box_332'; 333 'Box_323'; 334 'Box_334'; 335 'Box_335'; 336 'Box_336'; 337 'Box_337'; 338 'Box_338'; 339 'Box_339'; 340 'Box_340'; 341 'Box_341'; 342 'Box_342'; 343 'Box_343'; 344 'Box_344'; 345 'Box_345'; 346 'Box_346'; 347 'Box_347'; 348 'Box_348'; 349 'Box_349'; 350 'Box_350'; 351 'Box_351'; 352 'Box_352'; 353 'Box_353'; 354 'Box_354'; 355 'Box_355'; 356 'Box_356'; 357 'Box_357'; 358 'Box_358'; 359 'Box_359'; 360 'Box_360'; 361 'Box_361'; 362 'Box_362'; 363 'Box_363'; 364 'Box_364'; 365 'Box_365'; 366 'Box_366'; 367 'Box_367'; 368 'Box_368'; 369 'Box_369'; 370 'Box_370'; 371 'Box_371'; 372 'Box_372'; 373 'Box_373'; 374 'Box_374'; 375 'Box_375'; 376 'Box_376'; 377 'Box_377'; 378 'Box_378'; 379 'Box_379'; 380 'Box_380'; 381 'Box_381'; 382 'Box_382'; 383 'Box_383'; 384 'Box_384'; 385 'Box_385'; 386 'Box_386'; 387 'Box_387'; 388 'Box_388'; 389 'Box_389'; 390 'Box_390'; 391 'Box_391'; 392 'Box_392'; 393 'Box_393'; 394 'Box_394'; 395 'Box_395'; 396 'Box_396'; 397 'Box_397'; 398 'Box_398'; 399 'Box_399'; 400 'Box_400'; 401 'Box_401'; 402 'Box_402'; 403 'Box_403'; 404 'Box_404'; 405 'Box_405'; 406 'Box_406'; 407 'Box_407'; 408 'Box_408'; 409 'Box_409'; 410 'Box_410'; 411 'Box_411'; 412 'Box_412'; 413 'Box_413'; 414 'Box_414'; 415 'Box_415'; 416 'Box_416'; 417 'Box_417'; 418 'Box_418'; 419 'Box_419'; 420 'Box_420'; 421 'Box_421'; 422 'Box_422'; 423 'Box_423'; 424 'Box_424'; 425 'Box_425'; 426 'Box_426'; 427 'Box_427'; 428 'Box_428'; 429 'Box_429'; 430 'Box_430'; 431 'Box_431'; 432 'Box_432'; 433 'Box_433'; 434 'Box_434'; 435 'Box_435'; 436 'Box_436'; 437 'Box_437'; 438 'Box_438'; 439 'Box_439'; 440 'Box_440'; 441 'Box_441'; 442 'Box_442'; 443 'Box_443'; 444 'Box_444'; 445 'Box_445'; 446 'Box_446'; 447 'Box_447'; 448 'Box_448'; 449 'Box_449'; 450 'Box_450'; 451 'Box_451'; 452 'Box_452'; 453 'Box_453'; 454 'Box_454'; 455 'Box_455'; 456 'Box_456'; 457 'Box_457'; 458 'Box_458'; 459 'Box_459'; 460 'Box_460'; 461 'Box_461'; 462 'Box_462'; 463 'Box_463'; 464 'Box_464'; 465 'Box_465'; 466 'Box_466'; 467 'Box_467'; 468 'Box_468'; 469 'Box_469'; 470 'Box_470'; 471 'Box_471'; 472 'Box_472'; 473 'Box_473'; 474 'Box_474'; 475 'Box_475'; 476 'Box_476'; 477 'Box_477'; 478 'Box_478'; 479 'Box_479'; 480 'Box_480'; 481 'Box_481'; 482 'Box_482'; 483 'Box_483'; 484 'Box_484'; 485 'Box_485'; 486 'Box_486'; 487 'Box_487'; 488 'Box_488'; 489 'Box_489'; 490 'Box_490'; 491 'Box_491'; 492 'Box_492'; 493 'Box_493'; 494 'Box_494'; 495 'Box_495'; 496 'Box_496'; 497 'Box_497'; 498 'Box_498'; 499 'Box_499'; 500 'Box_500'; 501 'Box_501'; 502 'Box_502'; 503 'Box_503'; 504 'Box_504'; 505 'Box_505'; 506 'Box_506'; 507 'Box_507'; 508 'Box_508'; 509 'Box_509'; 510 'Box_510'; 511 'Box_511'; 512 'Box_512'; 513 'Box_513'; 514 'Box_514'; 515 'Box_515'; 516 'Box_516'; 517 'Box_517'; 518 'Box_518'; 519 'Box_519'; 520 'Box_520'; 521 'ช่องยานี้เต็มแล้ว'

text list "Zone_x 1.1": 0 '1'; 1 '8'; 2 '15'

text list "Zone_y1.5": 0 'E'; 1 'K'; 2 'Q'; 3 'W'

text list "Lisrt_Medicine2_1": 0 '1'; 1 '8'; 2 '15'

text list "Lisrt_Medicine2_2": 0 '2'; 1 '9'; 2 '16'

text list "Lisrt_Medicine2_3": 0 '3'; 1 '10'; 2 '17'

text list "Lisrt_Medicine2_5": 0 '5'; 1 '12'; 2 '19'

text list "Lisrt_Medicine2_4": 0 '4'; 1 '11'; 2 '18'

text list "Lisrt_Medicine_3": 0 'Zone_C'; 1 'Zone_I'; 2 'Zone_O'; 3 'Zone_U'

text list "Lisrt_Medicine_2": 0 'Zone_B'; 1 'Zone_H'; 2 'Zone_N'; 3 'Zone_T'; 4 'Zone_Z'

text list "Lisrt_Medicine_1": 0 'Zone_A'; 1 'Zone_G'; 2 'Zone_M'; 3 'Zone_S'; 4 'Zone_Y'

text list "Lisrt_Medicine_5": 0 'Zone_E'; 1 'Zone_K'; 2 'Zone_Q'; 3 'Zone_W'

text list "Lisrt_Medicine_4": 0 'Zone_D'; 1 'Zone_J'; 2 'Zone_P'; 3 'Zone_V'

text list "Lisrt_Medicine2_7": 0 '7'; 1 '14'

text list "Lisrt_Medicine_6": 0 'Zone_F'; 1 'Zone_L'; 2 'Zone_R'; 3 'Zone_X'

text list "Lisrt_Medicine2_6": 0 '6'; 1 '13'; 2 '20'

text list "SelectedMedicine": 0 'โปรดเลือกยา'; 1 'Lidocaine'; 2 'Bupivacaine'; 3 'Ropivacaine'; 4 'Procaine'; 5 'Benzocaine'; 6 'Tetracaine'; 7 'Propofol'; 8 'Ketamine'; 9 'Etomidate'; 10 'Thiopental'; 11 'Midazolam'; 12 'Diazepam'; 13 'Lorazepam'; 14 'Fentanyl'; 15 'Morphine'; 16 'Pethidine'; 17 'Tramadol'; 18 'Nalbuphine'; 19 'Remifentanil'; 20 'Succinylcholine'; 21 'Rocuronium'; 22 'Vecuronium'; 23 'Atracurium'; 24 'Cisatracurium'; 25 'Neostigmine'; 26 'Atropine'; 27 'Glycopyrrolate'; 28 'Epinephrine'; 29 'Norepinephrine'; 30 'Dopamine'; 31 'Dobutamine'; 32 'Phenylephrine'; 33 'Vasopressin'; 34 'Nitroglycerin'; 35 'Sodium nitroprusside'; 36 'Amiodarone'; 37 'Adenosine'; 38 'Verapamil'; 39 'Diltiazem'; 40 'Lidocaine'; 41 'Magnesium sulfate'; 42 'Calcium gluconate'; 43 'Sodium bicarbonate'; 44 'Potassium chloride'; 45 'Dextrose 50%'; 46 'Insulin regular'; 47 'Glucagon'; 48 'Hydrocortisone'; 49 'Dexamethasone'; 50 'Diphenhydramine'; 51 'Chlorpheniramine'; 52 'Salbutamol'; 53 'Ipratropium bromide'; 54 'Aminophylline'; 55 'Furosemide'; 56 'Mannitol'; 57 'Acetazolamide'; 58 'Tranexamic acid'; 59 'Vitamin K'; 60 'Protamine sulfate'; 61 'Naloxone'; 62 'Flumazenil'; 63 'Activated charcoal'; 64 'Acetylcysteine'; 65 'Deferoxamine'; 66 'Pralidoxime'; 67 'Atropine'; 68 'Methylene blue'; 69 'Succimer'; 70 'Digoxin immune fab'; 71 'Fomepizole'; 72 'Antivenom green pit viper'; 73 'Rabies immunoglobulin'; 74 'Tetanus immunoglobulin'; 75 'Human albumin'; 76 'Normal saline'; 77 'Heparin'; 78 'Enoxaparin'; 79 'Alteplase'; 80 'Streptokinase'; 81 'Urokinase'; 82 'Iohexol'; 83 'Iopamidol'; 84 'Iodixanol'; 85 'Gadopentetate dimeglumine'; 86 'Haloperidol'; 87 'Olanzapine'; 88 'Levetiracetam'; 89 'Phenytoin'; 90 'Sodium valproate'; 91 'Carbamazepine'; 92 'Phenobarbital'; 93 'Ketorolac'; 94 'Parecoxib'; 95 'Ondansetron'; 96 'Metoclopramide'; 97 'Granisetron'; 98 'Sugammadex'; 99 'Hydrocolloid dressing'; 100 'Paraffin gauze dressing'; 101 'Omeprazole'; 102 'Esomeprazole'; 103 'Pantoprazole'; 104 'Lansoprazole'; 105 'Dexlansoprazole'; 106 'Famotidine'; 107 'Cimetidine'; 108 'Sucralfate'; 109 'Aluminium hydroxide'; 110 'Magnesium hydroxide'; 111 'Simethicone'; 112 'Domperidone'; 113 'Metoclopramide'; 114 'Ondansetron'; 115 'Hyoscine butylbromide'; 116 'Bisacodyl'; 117 'Lactulose'; 118 'Senna'; 119 'ORS'; 120 'Loperamide'; 121 'Amlodipine'; 122 'Losartan'; 123 'Enalapril'; 124 'Captopril'; 125 'Lisinopril'; 126 'Hydrochlorothiazide'; 127 'Furosemide'; 128 'Spironolactone'; 129 'Atenolol'; 130 'Metoprolol'; 131 'Propranolol'; 132 'Carvedilol'; 133 'Digoxin'; 134 'Isosorbide dinitrate'; 135 'Nitroglycerin'; 136 'Aspirin'; 137 'Clopidogrel'; 138 'Warfarin'; 139 'Heparin'; 140 'Enoxaparin'; 141 'Simvastatin'; 142 'Atorvastatin'; 143 'Rosuvastatin'; 144 'Gemfibrozil'; 145 'Salbutamol'; 146 'Terbutaline'; 147 'Ipratropium bromide'; 148 'Tiotropium'; 149 'Budesonide'; 150 'Fluticasone'; 151 'Montelukast'; 152 'Theophylline'; 153 'Acetylcysteine'; 154 'Bromhexine'; 155 'Ambroxol'; 156 'Dextromethorphan'; 157 'Chlorpheniramine'; 158 'Loratadine'; 159 'Cetirizine'; 160 'Fexofenadine'; 161 'Paracetamol'; 162 'Ibuprofen'; 163 'Diclofenac'; 164 'Naproxen'; 165 'Celecoxib'; 166 'Tramadol'; 167 'Morphine'; 168 'Codeine'; 169 'Gabapentin'; 170 'Pregabalin'; 171 'Amitriptyline'; 172 'Nortriptyline'; 173 'Fluoxetine'; 174 'Sertraline'; 175 'Diazepam'; 176 'Lorazepam'; 177 'Alprazolam'; 178 'Clonazepam'; 179 'Phenytoin'; 180 'Sodium valproate'; 181 'Carbamazepine'; 182 'Levetiracetam'; 183 'Metformin'; 184 'Glibenclamide'; 185 'Gliclazide'; 186 'Pioglitazone'; 187 'Sitagliptin'; 188 'Insulin regular'; 189 'Insulin NPH'; 190 'Insulin glargine'; 191 'Levothyroxine'; 192 'Propylthiouracil'; 193 'Methimazole'; 194 'Prednisolone'; 195 'Dexamethasone'; 196 'Hydrocortisone'; 197 'Colchicine'; 198 'Allopurinol'; 199 'Febuxostat'; 200 'Calcium carbonate'; 201 'Vitamin B complex'; 202 'Vitamin C'; 203 'Ferrous fumarate'; 204 'Folic acid'; 205 'Cyanocobalamin'; 206 'Potassium chloride'; 207 'Sodium bicarbonate'; 208 'Calcium gluconate'; 209 'Magnesium sulfate'; 210 'Multivitamin'; 211 'Oral rehydration salt'; 212 'Baclofen'; 213 'Tizanidine'; 214 'Orphenadrine'; 215 'Meloxicam'; 216 'Piroxicam'; 217 'Etoricoxib'; 218 'Glucosamine'; 219 'Chondroitin sulfate'; 220 'Alendronate'; 221 'Amoxicillin'; 222 'Ampicillin'; 223 'Cloxacillin'; 224 'Dicloxacillin'; 225 'Penicillin V'; 226 'Benzathine penicillin G'; 227 'Piperacillin'; 228 'Ticarcillin'; 229 'Amoxicillin clavulanate'; 230 'Ampicillin sulbactam'; 231 'Cefalexin'; 232 'Cefadroxil'; 233 'Cefuroxime'; 234 'Cefixime'; 235 'Cefpodoxime'; 236 'Ceftriaxone'; 237 'Cefotaxime'; 238 'Ceftazidime'; 239 'Cefepime'; 240 'Cefoxitin'; 241 'Imipenem cilastatin'; 242 'Meropenem'; 243 'Ertapenem'; 244 'Aztreonam'; 245 'Vancomycin'; 246 'Teicoplanin'; 247 'Linezolid'; 248 'Daptomycin'; 249 'Gentamicin'; 250 'Amikacin'; 251 'Tobramycin'; 252 'Streptomycin'; 253 'Neomycin'; 254 'Erythromycin'; 255 'Clarithromycin'; 256 'Azithromycin'; 257 'Roxithromycin'; 258 'Clindamycin'; 259 'Lincomycin'; 260 'Doxycycline'; 261 'Tetracycline'; 262 'Minocycline'; 263 'Ciprofloxacin'; 264 'Levofloxacin'; 265 'Moxifloxacin'; 266 'Norfloxacin'; 267 'Ofloxacin'; 268 'Co-trimoxazole'; 269 'Sulfadiazine'; 270 'Sulfasalazine'; 271 'Metronidazole'; 272 'Tinidazole'; 273 'Nitrofurantoin'; 274 'Fosfomycin'; 275 'Rifampicin'; 276 'Isoniazid'; 277 'Ethambutol'; 278 'Pyrazinamide'; 279 'Ethionamide'; 280 'Cycloserine'; 281 'Fluconazole'; 282 'Itraconazole'; 283 'Ketoconazole'; 284 'Voriconazole'; 285 'Amphotericin B'; 286 'Nystatin'; 287 'Clotrimazole'; 288 'Miconazole'; 289 'Terbinafine'; 290 'Griseofulvin'; 291 'Acyclovir'; 292 'Valacyclovir'; 293 'Ganciclovir'; 294 'Oseltamivir'; 295 'Zanamivir'; 296 'Remdesivir'; 297 'Favipiravir'; 298 'Lamivudine'; 299 'Zidovudine'; 300 'Tenofovir'; 301 'Efavirenz'; 302 'Dolutegravir'; 303 'Nevirapine'; 304 'Lopinavir ritonavir'; 305 'Albendazole'; 306 'Mebendazole'; 307 'Ivermectin'; 308 'Praziquantel'; 309 'Pyrantel pamoate'; 310 'Diethylcarbamazine'; 311 'Chloroquine'; 312 'Primaquine'; 313 'Artesunate'; 314 'Artemether lumefantrine'; 315 'Quinine'; 316 'Dapsone'; 317 'Permethrin'; 318 'Benzyl benzoate'; 319 'Povidone iodine'; 320 'Chlorhexidine'; 321 'Colistin'; 322 'Caspofungin'; 323 'Bacitracin'; 324 'Fusidic acid'; 325 'Mupirocin'; 326 'Rabies vaccine'; 327 'Influenza vaccine'; 328 'Hepatitis B vaccine'; 329 'BCG vaccine'; 330 'DTP vaccine'; 331 'MMR vaccine'; 332 'JE vaccine'; 333 'HPV vaccine'; 334 'Varicella vaccine'; 335 'Pneumococcal vaccine'; 336 'Rotavirus vaccine'; 337 'COVID-19 vaccine'; 338 'Tetanus toxoid'; 339 'Rabies immunoglobulin'; 340 'Hepatitis B immunoglobulin'; 341 'Oxytocin'; 342 'Misoprostol'; 343 'Dinoprostone'; 344 'Methylergometrine'; 345 'Magnesium sulfate'; 346 'Nifedipine'; 347 'Terbutaline'; 348 'Ferrous fumarate'; 349 'Folic acid'; 350 'Calcium carbonate'; 351 'Ethinylestradiol'; 352 'Levonorgestrel'; 353 'Medroxyprogesterone'; 354 'Norethisterone'; 355 'Clomiphene citrate'; 356 'Letrozole'; 357 'Tamoxifen'; 358 'Anastrozole'; 359 'Exemestane'; 360 'Leuprolide'; 361 'Goserelin'; 362 'Finasteride'; 363 'Dutasteride'; 364 'Tamsulosin'; 365 'Alfuzosin'; 366 'Oxybutynin'; 367 'Tolterodine'; 368 'Solifenacin'; 369 'Mirabegron'; 370 'Potassium citrate'; 371 'Sodium bicarbonate'; 372 'Nitrofurantoin'; 373 'Fosfomycin'; 374 'Methotrexate'; 375 'Cyclophosphamide'; 376 'Ifosfamide'; 377 'Chlorambucil'; 378 'Melphalan'; 379 'Busulfan'; 380 'Cytarabine'; 381 'Fluorouracil'; 382 'Capecitabine'; 383 'Gemcitabine'; 384 'Doxorubicin'; 385 'Daunorubicin'; 386 'Epirubicin'; 387 'Bleomycin'; 388 'Vincristine'; 389 'Vinblastine'; 390 'Paclitaxel'; 391 'Docetaxel'; 392 'Cisplatin'; 393 'Carboplatin'; 394 'Oxaliplatin'; 395 'Irinotecan'; 396 'Etoposide'; 397 'Topotecan'; 398 'Hydroxyurea'; 399 'Mercaptopurine'; 400 'Thioguanine'; 401 'Imatinib'; 402 'Dasatinib'; 403 'Nilotinib'; 404 'Erlotinib'; 405 'Gefitinib'; 406 'Afatinib'; 407 'Sunitinib'; 408 'Sorafenib'; 409 'Lenvatinib'; 410 'Bevacizumab'; 411 'Trastuzumab'; 412 'Rituximab'; 413 'Pembrolizumab'; 414 'Nivolumab'; 415 'Ipilimumab'; 416 'Bicalutamide'; 417 'Flutamide'; 418 'Abiraterone'; 419 'Enzalutamide'; 420 'Megestrol acetate'; 421 'Zoledronic acid'; 422 'Pamidronate'; 423 'Calcitonin'; 424 'Denosumab'; 425 'Tacrolimus'; 426 'Cyclosporine'; 427 'Mycophenolate mofetil'; 428 'Azathioprine'; 429 'Sirolimus'; 430 'Everolimus'; 431 'Prednisolone'; 432 'Methylprednisolone'; 433 'Dexamethasone'; 434 'Basiliximab'; 435 'Anti-thymocyte globulin'; 436 'Interferon alfa'; 437 'Epoetin alfa'; 438 'Filgrastim'; 439 'Pegfilgrastim'; 440 'Romiplostim'; 441 'Thalidomide'; 442 'Lenalidomide'; 443 'Bortezomib'; 444 'Carfilzomib'; 445 'Daratumumab'; 446 'Mesna'; 447 'Leucovorin'; 448 'All-trans retinoic acid'; 449 'Arsenic trioxide'; 450 'Temozolomide'; 451 'Procarbazine'; 452 'Lomustine'; 453 'Carmustine'; 454 'Mitomycin C'; 455 'Actinomycin D'; 456 'Asparaginase'; 457 'Pegaspargase'; 458 'Brentuximab vedotin'; 459 'Olaparib'; 460 'Palbociclib'; 461 'Artificial tears'; 462 'Carboxy methylcellulose'; 463 'Hydroxypropyl methylcellulose'; 464 'Sodium hyaluronate'; 465 'Polyvinyl alcohol'; 466 'Timolol'; 467 'Betaxolol'; 468 'Brimonidine'; 469 'Dorzolamide'; 470 'Acetazolamide'; 471 'Latanoprost'; 472 'Travoprost'; 473 'Bimatoprost'; 474 'Pilocarpine'; 475 'Atropine'; 476 'Tropicamide'; 477 'Phenylephrine'; 478 'Ciprofloxacin'; 479 'Ofloxacin'; 480 'Moxifloxacin'; 481 'Tobramycin'; 482 'Gentamicin'; 483 'Chloramphenicol'; 484 'Fusidic acid'; 485 'Natamycin'; 486 'Acyclovir'; 487 'Prednisolone acetate'; 488 'Dexamethasone'; 489 'Fluorometholone'; 490 'Ketorolac'; 491 'Diclofenac'; 492 'Olopatadine'; 493 'Ketotifen'; 494 'Sodium cromoglycate'; 495 'Lubricating ointment'; 496 'Neomycin polymyxin B dexamethasone'; 497 'Oxymetazoline'; 498 'Xylometazoline'; 499 'Saline nasal spray'; 500 'Fluticasone'; 501 'Mometasone'; 502 'Budesonide'; 503 'Beclomethasone'; 504 'Azelastine'; 505 'Ipratropium bromide'; 506 'Menthol inhaler'; 507 'Carbamide peroxide'; 508 'Brinzolamide'; 509 'Ciprofloxacin'; 510 'Ofloxacin'; 511 'Neomycin polymyxin hydrocortisone'; 512 'Lidocaine'; 513 'Benzydamine'; 514 'Chlorhexidine'; 515 'Povidone iodine'; 516 'Nystatin'; 517 'Miconazole'; 518 'Triamcinolone acetonide'; 519 'Lidocaine viscous'; 520 'Sodium fluoride'

text list "X AXIS ( Horizontall )จัดเก็บ": 0 '0'; 1 '1353'; 2 '1270'; 3 '1187'; 4 '1104'; 5 '1021'; 6 '938'; 7 '855'; 8 '772'; 9 '689'; 10 '606'; 11 '523'; 12 '440'; 13 '357'; 14 '153'; 15 '70'; 16 '13'; 17 '96'; 18 '179'; 19 '262'; 20 '345'; 21 '428'; 22 '511'; 23 '594'; 24 '677'; 25 '760'; 26 '843'; 27 '1353'; 28 '1270'; 29 '1187'; 30 '1104'; 31 '1021'; 32 '938'; 33 '855'; 34 '772'; 35 '689'; 36 '606'; 37 '523'; 38 '440'; 39 '357'; 40 '153'; 41 '70'; 42 '13'; 43 '96'; 44 '179'; 45 '262'; 46 '345'; 47 '428'; 48 '511'; 49 '594'; 50 '677'; 51 '760'; 52 '843'; 53 '1353'; 54 '1270'; 55 '1187'; 56 '1104'; 57 '1021'; 58 '938'; 59 '855'; 60 '772'; 61 '689'; 62 '606'; 63 '523'; 64 '440'; 65 '357'; 66 '153'; 67 '70'; 68 '13'; 69 '96'; 70 '179'; 71 '262'; 72 '345'; 73 '428'; 74 '511'; 75 '594'; 76 '677'; 77 '760'; 78 '843'; 79 '1353'; 80 '1270'; 81 '1187'; 82 '1104'; 83 '1021'; 84 '938'; 85 '855'; 86 '772'; 87 '689'; 88 '606'; 89 '523'; 90 '440'; 91 '357'; 92 '153'; 93 '70'; 94 '13'; 95 '96'; 96 '179'; 97 '262'; 98 '345'; 99 '428'; 100 '511'; 101 '594'; 102 '677'; 103 '760'; 104 '843'; 105 '1353'; 106 '1270'; 107 '1187'; 108 '1104'; 109 '1021'; 110 '938'; 111 '855'; 112 '772'; 113 '689'; 114 '606'; 115 '523'; 116 '440'; 117 '357'; 118 '153'; 119 '70'; 120 '13'; 121 '96'; 122 '179'; 123 '262'; 124 '345'; 125 '428'; 126 '511'; 127 '594'; 128 '677'; 129 '760'; 130 '843'; 131 '1353'; 132 '1270'; 133 '1187'; 134 '1104'; 135 '1021'; 136 '938'; 137 '855'; 138 '772'; 139 '689'; 140 '606'; 141 '523'; 142 '440'; 143 '357'; 144 '153'; 145 '70'; 146 '13'; 147 '96'; 148 '179'; 149 '262'; 150 '345'; 151 '428'; 152 '511'; 153 '594'; 154 '677'; 155 '760'; 156 '843'; 157 '1353'; 158 '1270'; 159 '1187'; 160 '1104'; 161 '1021'; 162 '938'; 163 '855'; 164 '772'; 165 '689'; 166 '606'; 167 '523'; 168 '440'; 169 '357'; 170 '153'; 171 '70'; 172 '13'; 173 '96'; 174 '179'; 175 '262'; 176 '345'; 177 '428'; 178 '511'; 179 '594'; 180 '677'; 181 '760'; 182 '843'; 183 '1353'; 184 '1270'; 185 '1187'; 186 '1104'; 187 '1021'; 188 '938'; 189 '855'; 190 '772'; 191 '689'; 192 '606'; 193 '523'; 194 '440'; 195 '357'; 196 '153'; 197 '70'; 198 '13'; 199 '96'; 200 '179'; 201 '262'; 202 '345'; 203 '428'; 204 '511'; 205 '594'; 206 '677'; 207 '760'; 208 '843'; 209 '1353'; 210 '1270'; 211 '1187'; 212 '1104'; 213 '1021'; 214 '938'; 215 '855'; 216 '772'; 217 '689'; 218 '606'; 219 '523'; 220 '440'; 221 '357'; 222 '153'; 223 '70'; 224 '13'; 225 '96'; 226 '179'; 227 '262'; 228 '345'; 229 '428'; 230 '511'; 231 '594'; 232 '677'; 233 '760'; 234 '843'; 235 '1353'; 236 '1270'; 237 '1187'; 238 '1104'; 239 '1021'; 240 '938'; 241 '855'; 242 '772'; 243 '689'; 244 '606'; 245 '523'; 246 '440'; 247 '357'; 248 '153'; 249 '70'; 250 '13'; 251 '96'; 252 '179'; 253 '262'; 254 '345'; 255 '428'; 256 '511'; 257 '594'; 258 '677'; 259 '760'; 260 '843'; 261 '1353'; 262 '1270'; 263 '1187'; 264 '1104'; 265 '1021'; 266 '938'; 267 '855'; 268 '772'; 269 '689'; 270 '606'; 271 '523'; 272 '440'; 273 '357'; 274 '153'; 275 '70'; 276 '13'; 277 '96'; 278 '179'; 279 '262'; 280 '345'; 281 '428'; 282 '511'; 283 '594'; 284 '677'; 285 '760'; 286 '843'; 287 '1353'; 288 '1270'; 289 '1187'; 290 '1104'; 291 '1021'; 292 '938'; 293 '855'; 294 '772'; 295 '689'; 296 '606'; 297 '523'; 298 '440'; 299 '357'; 300 '153'; 301 '70'; 302 '13'; 303 '96'; 304 '179'; 305 '262'; 306 '345'; 307 '428'; 308 '511'; 309 '594'; 310 '677'; 311 '760'; 312 '843'; 313 '1353'; 314 '1270'; 315 '1187'; 316 '1104'; 317 '1021'; 318 '938'; 319 '855'; 320 '772'; 321 '689'; 322 '606'; 323 '523'; 324 '440'; 325 '357'; 326 '153'; 327 '70'; 328 '13'; 329 '96'; 330 '179'; 331 '262'; 332 '345'; 333 '428'; 334 '511'; 335 '594'; 336 '677'; 337 '760'; 338 '843'; 339 '1353'; 340 '1270'; 341 '1187'; 342 '1104'; 343 '1021'; 344 '938'; 345 '855'; 346 '772'; 347 '689'; 348 '606'; 349 '523'; 350 '440'; 351 '357'; 352 '153'; 353 '70'; 354 '13'; 355 '96'; 356 '179'; 357 '262'; 358 '345'; 359 '428'; 360 '511'; 361 '594'; 362 '677'; 363 '760'; 364 '843'; 365 '1353'; 366 '1270'; 367 '1187'; 368 '1104'; 369 '1021'; 370 '938'; 371 '855'; 372 '772'; 373 '689'; 374 '606'; 375 '523'; 376 '440'; 377 '357'; 378 '153'; 379 '70'; 380 '13'; 381 '96'; 382 '179'; 383 '262'; 384 '345'; 385 '428'; 386 '511'; 387 '594'; 388 '677'; 389 '760'; 390 '843'; 391 '1353'; 392 '1270'; 393 '1187'; 394 '1104'; 395 '1021'; 396 '938'; 397 '855'; 398 '772'; 399 '689'; 400 '606'; 401 '523'; 402 '440'; 403 '357'; 404 '153'; 405 '70'; 406 '13'; 407 '96'; 408 '179'; 409 '262'; 410 '345'; 411 '428'; 412 '511'; 413 '594'; 414 '677'; 415 '760'; 416 '843'; 417 '1353'; 418 '1270'; 419 '1187'; 420 '1104'; 421 '1021'; 422 '938'; 423 '855'; 424 '772'; 425 '689'; 426 '606'; 427 '523'; 428 '440'; 429 '357'; 430 '153'; 431 '70'; 432 '13'; 433 '96'; 434 '179'; 435 '262'; 436 '345'; 437 '428'; 438 '511'; 439 '594'; 440 '677'; 441 '760'; 442 '843'; 443 '1353'; 444 '1270'; 445 '1187'; 446 '1104'; 447 '1021'; 448 '938'; 449 '855'; 450 '772'; 451 '689'; 452 '606'; 453 '523'; 454 '440'; 455 '357'; 456 '153'; 457 '70'; 458 '13'; 459 '96'; 460 '179'; 461 '262'; 462 '345'; 463 '428'; 464 '511'; 465 '594'; 466 '677'; 467 '760'; 468 '843'; 469 '1353'; 470 '1270'; 471 '1187'; 472 '1104'; 473 '1021'; 474 '938'; 475 '855'; 476 '772'; 477 '689'; 478 '606'; 479 '523'; 480 '440'; 481 '357'; 482 '153'; 483 '70'; 484 '13'; 485 '96'; 486 '179'; 487 '262'; 488 '345'; 489 '428'; 490 '511'; 491 '594'; 492 '677'; 493 '760'; 494 '843'

text list "Y AXIS ( Verticall )จัดเก็บ": 0 '0'; 1..26 '1466'; 27..52 '1371.00'; 53..78 '1276.00'; 79..104 '1181.00'; 105..130 '1086.00'; 131..156 '991.00'; 157..182 '896.00'; 183..208 '801.00'; 209..234 '706.00'; 235..260 '611.00'; 261..286 '516.00'; 287..312 '421.00'; 313..338 '326.00'; 339..364 '231.00'; 365..390 '136.00'; 391..416 '41.00'; 417..442 '-54.00'; 443..468 '-149.00'; 469..494 '-244.00'

text list "poperty": 0 'STOP'; 1 'RUNNING'

text list "EncoderแกนY (เบิกจ่าย)": 0 '0'; 1..26 '27619'; 27..52 '23934'; 53..78 '20249'; 79..104 '16564'; 105..130 '12879'; 131..156 '9194'; 157..182 '5509'; 183..208 '1824'; 209..234 '1861'; 235..260 '5546'; 261..286 '9231'; 287..312 '12916'; 313..338 '16601'; 339..364 '20286'; 365..390 '23971'; 391..416 '27656'; 417..442 '31341'; 443..468 '35026'; 469..494 '38711'

text list "EncoderแกนX (จัดเก็บ)": 0 '0'; 1 '52483'; 2 '49263'; 3 '46043'; 4 '42823'; 5 '39603'; 6 '36383'; 7 '33163'; 8 '29943'; 9 '26723'; 10 '23503'; 11 '20283'; 12 '17063'; 13 '13843'; 14 '5935'; 15 '2715'; 16 '505'; 17 '3725'; 18 '6945'; 19 '10165'; 20 '13385'; 21 '16605'; 22 '19825'; 23 '23045'; 24 '26265'; 25 '29485'; 26 '32705'; 27 '52483'; 28 '49263'; 29 '46043'; 30 '42823'; 31 '39603'; 32 '36383'; 33 '33163'; 34 '29943'; 35 '26723'; 36 '23503'; 37 '20283'; 38 '17063'; 39 '13843'; 40 '5935'; 41 '2715'; 42 '505'; 43 '3725'; 44 '6945'; 45 '10165'; 46 '13385'; 47 '16605'; 48 '19825'; 49 '23045'; 50 '26265'; 51 '29485'; 52 '32705'; 53 '52483'; 54 '49263'; 55 '46043'; 56 '42823'; 57 '39603'; 58 '36383'; 59 '33163'; 60 '29943'; 61 '26723'; 62 '23503'; 63 '20283'; 64 '17063'; 65 '13843'; 66 '5935'; 67 '2715'; 68 '505'; 69 '3725'; 70 '6945'; 71 '10165'; 72 '13385'; 73 '16605'; 74 '19825'; 75 '23045'; 76 '26265'; 77 '29485'; 78 '32705'; 79 '52483'; 80 '49263'; 81 '46043'; 82 '42823'; 83 '39603'; 84 '36383'; 85 '33163'; 86 '29943'; 87 '26723'; 88 '23503'; 89 '20283'; 90 '17063'; 91 '13843'; 92 '5935'; 93 '2715'; 94 '505'; 95 '3725'; 96 '6945'; 97 '10165'; 98 '13385'; 99 '16605'; 100 '19825'; 101 '23045'; 102 '26265'; 103 '29485'; 104 '32705'; 105 '52483'; 106 '49263'; 107 '46043'; 108 '42823'; 109 '39603'; 110 '36383'; 111 '33163'; 112 '29943'; 113 '26723'; 114 '23503'; 115 '20283'; 116 '17063'; 117 '13843'; 118 '5935'; 119 '2715'; 120 '505'; 121 '3725'; 122 '6945'; 123 '10165'; 124 '13385'; 125 '16605'; 126 '19825'; 127 '23045'; 128 '26265'; 129 '29485'; 130 '32705'; 131 '52483'; 132 '49263'; 133 '46043'; 134 '42823'; 135 '39603'; 136 '36383'; 137 '33163'; 138 '29943'; 139 '26723'; 140 '23503'; 141 '20283'; 142 '17063'; 143 '13843'; 144 '5935'; 145 '2715'; 146 '505'; 147 '3725'; 148 '6945'; 149 '10165'; 150 '13385'; 151 '16605'; 152 '19825'; 153 '23045'; 154 '26265'; 155 '29485'; 156 '32705'; 157 '52483'; 158 '49263'; 159 '46043'; 160 '42823'; 161 '39603'; 162 '36383'; 163 '33163'; 164 '29943'; 165 '26723'; 166 '23503'; 167 '20283'; 168 '17063'; 169 '13843'; 170 '5935'; 171 '2715'; 172 '505'; 173 '3725'; 174 '6945'; 175 '10165'; 176 '13385'; 177 '16605'; 178 '19825'; 179 '23045'; 180 '26265'; 181 '29485'; 182 '32705'; 183 '52483'; 184 '49263'; 185 '46043'; 186 '42823'; 187 '39603'; 188 '36383'; 189 '33163'; 190 '29943'; 191 '26723'; 192 '23503'; 193 '20283'; 194 '17063'; 195 '13843'; 196 '5935'; 197 '2715'; 198 '505'; 199 '3725'; 200 '6945'; 201 '10165'; 202 '13385'; 203 '16605'; 204 '19825'; 205 '23045'; 206 '26265'; 207 '29485'; 208 '32705'; 209 '52483'; 210 '49263'; 211 '46043'; 212 '42823'; 213 '39603'; 214 '36383'; 215 '33163'; 216 '29943'; 217 '26723'; 218 '23503'; 219 '20283'; 220 '17063'; 221 '13843'; 222 '5935'; 223 '2715'; 224 '505'; 225 '3725'; 226 '6945'; 227 '10165'; 228 '13385'; 229 '16605'; 230 '19825'; 231 '23045'; 232 '26265'; 233 '29485'; 234 '32705'; 235 '52483'; 236 '49263'; 237 '46043'; 238 '42823'; 239 '39603'; 240 '36383'; 241 '33163'; 242 '29943'; 243 '26723'; 244 '23503'; 245 '20283'; 246 '17063'; 247 '13843'; 248 '5935'; 249 '2715'; 250 '505'; 251 '3725'; 252 '6945'; 253 '10165'; 254 '13385'; 255 '16605'; 256 '19825'; 257 '23045'; 258 '26265'; 259 '29485'; 260 '32705'; 261 '52483'; 262 '49263'; 263 '46043'; 264 '42823'; 265 '39603'; 266 '36383'; 267 '33163'; 268 '29943'; 269 '26723'; 270 '23503'; 271 '20283'; 272 '17063'; 273 '13843'; 274 '5935'; 275 '2715'; 276 '505'; 277 '3725'; 278 '6945'; 279 '10165'; 280 '13385'; 281 '16605'; 282 '19825'; 283 '23045'; 284 '26265'; 285 '29485'; 286 '32705'; 287 '52483'; 288 '49263'; 289 '46043'; 290 '42823'; 291 '39603'; 292 '36383'; 293 '33163'; 294 '29943'; 295 '26723'; 296 '23503'; 297 '20283'; 298 '17063'; 299 '13843'; 300 '5935'; 301 '2715'; 302 '505'; 303 '3725'; 304 '6945'; 305 '10165'; 306 '13385'; 307 '16605'; 308 '19825'; 309 '23045'; 310 '26265'; 311 '29485'; 312 '32705'; 313 '52483'; 314 '49263'; 315 '46043'; 316 '42823'; 317 '39603'; 318 '36383'; 319 '33163'; 320 '29943'; 321 '26723'; 322 '23503'; 323 '20283'; 324 '17063'; 325 '13843'; 326 '5935'; 327 '2715'; 328 '505'; 329 '3725'; 330 '6945'; 331 '10165'; 332 '13385'; 333 '16605'; 334 '19825'; 335 '23045'; 336 '26265'; 337 '29485'; 338 '32705'; 339 '52483'; 340 '49263'; 341 '46043'; 342 '42823'; 343 '39603'; 344 '36383'; 345 '33163'; 346 '29943'; 347 '26723'; 348 '23503'; 349 '20283'; 350 '17063'; 351 '13843'; 352 '5935'; 353 '2715'; 354 '505'; 355 '3725'; 356 '6945'; 357 '10165'; 358 '13385'; 359 '16605'; 360 '19825'; 361 '23045'; 362 '26265'; 363 '29485'; 364 '32705'; 365 '52483'; 366 '49263'; 367 '46043'; 368 '42823'; 369 '39603'; 370 '36383'; 371 '33163'; 372 '29943'; 373 '26723'; 374 '23503'; 375 '20283'; 376 '17063'; 377 '13843'; 378 '5935'; 379 '2715'; 380 '505'; 381 '3725'; 382 '6945'; 383 '10165'; 384 '13385'; 385 '16605'; 386 '19825'; 387 '23045'; 388 '26265'; 389 '29485'; 390 '32705'; 391 '52483'; 392 '49263'; 393 '46043'; 394 '42823'; 395 '39603'; 396 '36383'; 397 '33163'; 398 '29943'; 399 '26723'; 400 '23503'; 401 '20283'; 402 '17063'; 403 '13843'; 404 '5935'; 405 '2715'; 406 '505'; 407 '3725'; 408 '6945'; 409 '10165'; 410 '13385'; 411 '16605'; 412 '19825'; 413 '23045'; 414 '26265'; 415 '29485'; 416 '32705'; 417 '52483'; 418 '49263'; 419 '46043'; 420 '42823'; 421 '39603'; 422 '36383'; 423 '33163'; 424 '29943'; 425 '26723'; 426 '23503'; 427 '20283'; 428 '17063'; 429 '13843'; 430 '5935'; 431 '2715'; 432 '505'; 433 '3725'; 434 '6945'; 435 '10165'; 436 '13385'; 437 '16605'; 438 '19825'; 439 '23045'; 440 '26265'; 441 '29485'; 442 '32705'; 443 '52483'; 444 '49263'; 445 '46043'; 446 '42823'; 447 '39603'; 448 '36383'; 449 '33163'; 450 '29943'; 451 '26723'; 452 '23503'; 453 '20283'; 454 '17063'; 455 '13843'; 456 '5935'; 457 '2715'; 458 '505'; 459 '3725'; 460 '6945'; 461 '10165'; 462 '13385'; 463 '16605'; 464 '19825'; 465 '23045'; 466 '26265'; 467 '29485'; 468 '32705'; 469 '52483'; 470 '49263'; 471 '46043'; 472 '42823'; 473 '39603'; 474 '36383'; 475 '33163'; 476 '29943'; 477 '26723'; 478 '23503'; 479 '20283'; 480 '17063'; 481 '13843'; 482 '5935'; 483 '2715'; 484 '505'; 485 '3725'; 486 '6945'; 487 '10165'; 488 '13385'; 489 '16605'; 490 '19825'; 491 '23045'; 492 '26265'; 493 '29485'; 494 '32705'

text list "EncoderแกนY (จัดเก็บ)": 0 '0'; 1..26 '56866'; 27..52 '53181'; 53..78 '49496'; 79..104 '45811'; 105..130 '42126'; 131..156 '38441'; 157..182 '34756'; 183..208 '31071'; 209..234 '27386'; 235..260 '23701'; 261..286 '20016'; 287..312 '16331'; 313..338 '12646'; 339..364 '8961'; 365..390 '5276'; 391..416 '1591'; 417..442 '2094'; 443..468 '5779'; 469..494 '9464'

text list "X AXIS ( Horizontall )เบิกจ่าย": 0 '0'; 1 '153'; 2 '236'; 3 '319'; 4 '402'; 5 '485'; 6 '568'; 7 '651'; 8 '734'; 9 '817'; 10 '900'; 11 '983'; 12 '1066'; 13 '1149'; 14 '1353'; 15 '1436'; 16 '1519'; 17 '1602'; 18 '1685'; 19 '1768'; 20 '1851'; 21 '1934'; 22 '2017'; 23 '2100'; 24 '2183'; 25 '2266'; 26 '2349'; 27 '153'; 28 '236'; 29 '319'; 30 '402'; 31 '485'; 32 '568'; 33 '651'; 34 '734'; 35 '817'; 36 '900'; 37 '983'; 38 '1066'; 39 '1149'; 40 '1353'; 41 '1436'; 42 '1519'; 43 '1602'; 44 '1685'; 45 '1768'; 46 '1851'; 47 '1934'; 48 '2017'; 49 '2100'; 50 '2183'; 51 '2266'; 52 '2349'; 53 '153'; 54 '236'; 55 '319'; 56 '402'; 57 '485'; 58 '568'; 59 '651'; 60 '734'; 61 '817'; 62 '900'; 63 '983'; 64 '1066'; 65 '1149'; 66 '1353'; 67 '1436'; 68 '1519'; 69 '1602'; 70 '1685'; 71 '1768'; 72 '1851'; 73 '1934'; 74 '2017'; 75 '2100'; 76 '2183'; 77 '2266'; 78 '2349'; 79 '153'; 80 '236'; 81 '319'; 82 '402'; 83 '485'; 84 '568'; 85 '651'; 86 '734'; 87 '817'; 88 '900'; 89 '983'; 90 '1066'; 91 '1149'; 92 '1353'; 93 '1436'; 94 '1519'; 95 '1602'; 96 '1685'; 97 '1768'; 98 '1851'; 99 '1934'; 100 '2017'; 101 '2100'; 102 '2183'; 103 '2266'; 104 '2349'; 105 '153'; 106 '236'; 107 '319'; 108 '402'; 109 '485'; 110 '568'; 111 '651'; 112 '734'; 113 '817'; 114 '900'; 115 '983'; 116 '1066'; 117 '1149'; 118 '1353'; 119 '1436'; 120 '1519'; 121 '1602'; 122 '1685'; 123 '1768'; 124 '1851'; 125 '1934'; 126 '2017'; 127 '2100'; 128 '2183'; 129 '2266'; 130 '2349'; 131 '153'; 132 '236'; 133 '319'; 134 '402'; 135 '485'; 136 '568'; 137 '651'; 138 '734'; 139 '817'; 140 '900'; 141 '983'; 142 '1066'; 143 '1149'; 144 '1353'; 145 '1436'; 146 '1519'; 147 '1602'; 148 '1685'; 149 '1768'; 150 '1851'; 151 '1934'; 152 '2017'; 153 '2100'; 154 '2183'; 155 '2266'; 156 '2349'; 157 '153'; 158 '236'; 159 '319'; 160 '402'; 161 '485'; 162 '568'; 163 '651'; 164 '734'; 165 '817'; 166 '900'; 167 '983'; 168 '1066'; 169 '1149'; 170 '1353'; 171 '1436'; 172 '1519'; 173 '1602'; 174 '1685'; 175 '1768'; 176 '1851'; 177 '1934'; 178 '2017'; 179 '2100'; 180 '2183'; 181 '2266'; 182 '2349'; 183 '153'; 184 '236'; 185 '319'; 186 '402'; 187 '485'; 188 '568'; 189 '651'; 190 '734'; 191 '817'; 192 '900'; 193 '983'; 194 '1066'; 195 '1149'; 196 '1353'; 197 '1436'; 198 '1519'; 199 '1602'; 200 '1685'; 201 '1768'; 202 '1851'; 203 '1934'; 204 '2017'; 205 '2100'; 206 '2183'; 207 '2266'; 208 '2349'; 209 '153'; 210 '236'; 211 '319'; 212 '402'; 213 '485'; 214 '568'; 215 '651'; 216 '734'; 217 '817'; 218 '900'; 219 '983'; 220 '1066'; 221 '1149'; 222 '1353'; 223 '1436'; 224 '1519'; 225 '1602'; 226 '1685'; 227 '1768'; 228 '1851'; 229 '1934'; 230 '2017'; 231 '2100'; 232 '2183'; 233 '2266'; 234 '2349'; 235 '153'; 236 '236'; 237 '319'; 238 '402'; 239 '485'; 240 '568'; 241 '651'; 242 '734'; 243 '817'; 244 '900'; 245 '983'; 246 '1066'; 247 '1149'; 248 '1353'; 249 '1436'; 250 '1519'; 251 '1602'; 252 '1685'; 253 '1768'; 254 '1851'; 255 '1934'; 256 '2017'; 257 '2100'; 258 '2183'; 259 '2266'; 260 '2349'; 261 '153'; 262 '236'; 263 '319'; 264 '402'; 265 '485'; 266 '568'; 267 '651'; 268 '734'; 269 '817'; 270 '900'; 271 '983'; 272 '1066'; 273 '1149'; 274 '1353'; 275 '1436'; 276 '1519'; 277 '1602'; 278 '1685'; 279 '1768'; 280 '1851'; 281 '1934'; 282 '2017'; 283 '2100'; 284 '2183'; 285 '2266'; 286 '2349'; 287 '153'; 288 '236'; 289 '319'; 290 '402'; 291 '485'; 292 '568'; 293 '651'; 294 '734'; 295 '817'; 296 '900'; 297 '983'; 298 '1066'; 299 '1149'; 300 '1353'; 301 '1436'; 302 '1519'; 303 '1602'; 304 '1685'; 305 '1768'; 306 '1851'; 307 '1934'; 308 '2017'; 309 '2100'; 310 '2183'; 311 '2266'; 312 '2349'; 313 '153'; 314 '236'; 315 '319'; 316 '402'; 317 '485'; 318 '568'; 319 '651'; 320 '734'; 321 '817'; 322 '900'; 323 '983'; 324 '1066'; 325 '1149'; 326 '1353'; 327 '1436'; 328 '1519'; 329 '1602'; 330 '1685'; 331 '1768'; 332 '1851'; 333 '1934'; 334 '2017'; 335 '2100'; 336 '2183'; 337 '2266'; 338 '2349'; 339 '153'; 340 '236'; 341 '319'; 342 '402'; 343 '485'; 344 '568'; 345 '651'; 346 '734'; 347 '817'; 348 '900'; 349 '983'; 350 '1066'; 351 '1149'; 352 '1353'; 353 '1436'; 354 '1519'; 355 '1602'; 356 '1685'; 357 '1768'; 358 '1851'; 359 '1934'; 360 '2017'; 361 '2100'; 362 '2183'; 363 '2266'; 364 '2349'; 365 '153'; 366 '236'; 367 '319'; 368 '402'; 369 '485'; 370 '568'; 371 '651'; 372 '734'; 373 '817'; 374 '900'; 375 '983'; 376 '1066'; 377 '1149'; 378 '1353'; 379 '1436'; 380 '1519'; 381 '1602'; 382 '1685'; 383 '1768'; 384 '1851'; 385 '1934'; 386 '2017'; 387 '2100'; 388 '2183'; 389 '2266'; 390 '2349'; 391 '153'; 392 '236'; 393 '319'; 394 '402'; 395 '485'; 396 '568'; 397 '651'; 398 '734'; 399 '817'; 400 '900'; 401 '983'; 402 '1066'; 403 '1149'; 404 '1353'; 405 '1436'; 406 '1519'; 407 '1602'; 408 '1685'; 409 '1768'; 410 '1851'; 411 '1934'; 412 '2017'; 413 '2100'; 414 '2183'; 415 '2266'; 416 '2349'; 417 '153'; 418 '236'; 419 '319'; 420 '402'; 421 '485'; 422 '568'; 423 '651'; 424 '734'; 425 '817'; 426 '900'; 427 '983'; 428 '1066'; 429 '1149'; 430 '1353'; 431 '1436'; 432 '1519'; 433 '1602'; 434 '1685'; 435 '1768'; 436 '1851'; 437 '1934'; 438 '2017'; 439 '2100'; 440 '2183'; 441 '2266'; 442 '2349'; 443 '153'; 444 '236'; 445 '319'; 446 '402'; 447 '485'; 448 '568'; 449 '651'; 450 '734'; 451 '817'; 452 '900'; 453 '983'; 454 '1066'; 455 '1149'; 456 '1353'; 457 '1436'; 458 '1519'; 459 '1602'; 460 '1685'; 461 '1768'; 462 '1851'; 463 '1934'; 464 '2017'; 465 '2100'; 466 '2183'; 467 '2266'; 468 '2349'; 469 '153'; 470 '236'; 471 '319'; 472 '402'; 473 '485'; 474 '568'; 475 '651'; 476 '734'; 477 '817'; 478 '900'; 479 '983'; 480 '1066'; 481 '1149'; 482 '1353'; 483 '1436'; 484 '1519'; 485 '1602'; 486 '1685'; 487 '1768'; 488 '1851'; 489 '1934'; 490 '2017'; 491 '2100'; 492 '2183'; 493 '2266'; 494 '2349'

text list "Y AXIS ( Verticall )เบิกจ่่าย": 0 '0'; 1..26 '712'; 27..52 '617'; 53..78 '522'; 79..104 '427'; 105..130 '332'; 131..156 '237'; 157..182 '142'; 183..208 '47'; 209..234 '-48'; 235..260 '-143'; 261..286 '-238'; 287..312 '-333'; 313..338 '-428'; 339..364 '-523'; 365..390 '-618'; 391..416 '-713'; 417..442 '-808'; 443..468 '-903'; 469..494 '-998'

text list "จำนวนกล่องยาที่เลือกหน้า Or": 0 '0'; 1 '1'

